(* IEC 61131-3 sources: daoli-st-library/DL_Device (part 3) *)

(* ---- FB_DL_HydraulicPowerUnit.st ---- *)
(*==============================================================================
 * 组件名称 (Component)  : FB_DL_HydraulicPowerUnit
 * 所属子库 (Sublibrary) : DL_Device
 * 当前版本 (Version)    : 1.0.0
 * 兼容性   (Platform)   : CODESYS 3.5+ / TwinCAT 3 / 汇川 InoProShop / 施耐德 Machine Expert
 *                         仅依赖 Standard.library（TON / R_TRIG），零厂商私有库
 * 功能描述 (Function)   : 液压动力单元（HPU）顺控：bStart 上升沿先查油温/油位
 *                         联锁（先于电机判据，规格指定），通过后启动电机升压；
 *                         压力达 fPressSwMpa 开卸荷阀，压力回落至 (fPressSwMpa
 *                         − 0.5 MPa) 关卸荷阀（±0.5 MPa 回差顺控，规格指定）；
 *                         电机启停切换设最小间隔互锁 tMinSw（切换后 tMinSw 内
 *                         禁再次切换）。运行中油温超限/油位低于下限/压力非有限
 *                         → 停电机锁存故障（安全侧优先）。
 * 接口     (Interface)  : 输入 bStart 启动命令（上升沿触发，FALSE 停机）、fPressMpa
 *                         压力实测 [MPa]、fOilTempC 油温实测 [℃]、fOilLevelPct
 *                         油位实测 [%]、fPressSwMpa 卸荷切换阈（域 > 0.5）、
 *                         fTempMaxC 油温联锁上限（域 > 0）、fLvlMinPct 油位联锁
 *                         下限（域 > 0 且 < 100）、tMinSw 电机切换最小间隔、
 *                         bReset 复位；输出 bMotor 电机命令、bUnload 卸荷阀
 *                         命令、ePhase 五态相位、eErrCode 错误码、bError 故障
 *                         标志。
 * 边界     (Boundary)   : ① **属主边界（写死）：本件只出电机/卸荷阀命令，不驱动
 *                         接触器/阀线圈本体**；执行器驱动归 IO 映射层（DOL 电机
 *                         包装归 `FB_DL_DolMotor`）。
 *                         ② 五态 CASE + ELSE 兜底（R6）；tonMinSw IN 挂切换
 *                         互锁窗本身（切换后置互锁、到时解除），三 TON 两沿段 0
 *                         无条件调用（R7）。
 *                         ③ 联锁先于电机判据：启动沿先查油温/油位，联锁不过
 *                         不入启动相并置信息码 eInterlock（不锁存故障，联锁
 *                         为常态门槛）；运行中联锁破约才锁存故障 eTempHigh/
 *                         eLvlLow（归因唯一，R190）。
 *                         ④ 回差口径：开阀阈 fPressSwMpa，关阀阈 fPressSwMpa
 *                         − DL_HPU_DBAND(0.5 MPa)，组态闸保证 fPressSwMpa >
 *                         0.5（关阀阈恒正）。
 *                         ⑤ 电机切换互锁：每次 bMotor 电平变化后 _bSwBlock 置
 *                         位，tonMinSw 到时解除；互锁期内启动/停止命令一律
 *                         拒绝（拒动安全侧）。
 *                         ⑥ 压力非有限（R79 双判）运行中 → 停电机锁存
 *                         ePressBad（不可判即安全侧停机）。
 *                         ⑦ 零全局耦合（无 GVL / VAR_EXTERNAL / 物理地址）。
 * 分工声明 (Scope)      : 与 `FB_DL_DolMotor` 分工：电机直启包装归那件、HPU 工艺
 *                         顺控归本件；与 `FB_DL_MinOnOffGuard` 分工：通用最小
 *                         启停保护归那件，本件互锁为切换间隔专用语义。
 * 来源标签 (Source Tag) : 自研线（卸荷回差顺控为公开液压系统控制实践 clean-room）
 * 码表     (Codes)      : 本件不占用任何全局数字码位。出口为 BOOL 命令组 +
 *                         ENUM 相位/错误码；数字码位待主控收口阶段统一派号。
 * 红线自检 (Redline)    : R1 ✓ 零 GVL/VAR_EXTERNAL ｜ R2 ✓ 零 %I/%Q/%M ｜ R3 ✓ 纯 IEC 61131-3
 *                         R4 ✓ 联锁前置 + 回差 + 切换互锁 + 非有限安全停机
 *                         ｜ R5 ✓ 声明逐行同行双语注释
 *                         R6 ✓ 五态 CASE 含 ELSE ｜ R7 ✓ 三 TON 两 R_TRIG 段 0 无条件刷新
 * 修订历史 (Revision)   : 2026-11-20  v1.0.0  R50 首版（批次 4 · 序号 18）
 * 验收向量 (Acceptance) : ① 油位 25%（下限 30%）时启动沿 → 不入启动相，
 *                         eErrCode=eInterlock，bMotor=FALSE；② 正常启动，
 *                         压力升至 16.2 MPa（阈 16.0）→ bUnload=TRUE；回落至
 *                         15.4 MPa（< 16.0−0.5=15.5）→ bUnload=FALSE；③ 运行
 *                         中油温 65 ℃（上限 60）→ 停电机锁存 eTempHigh；
 *                         ④ 停机后 2s 内再启动（tMinSw=10S）→ 拒动（互锁）。
 *==============================================================================*)

(*-----------------------------------------------------------------------------
 * 枚举: E_DL_HpuPhase（HPU 相位，全库唯一属主本文件）
 *----------------------------------------------------------------------------*)
TYPE E_DL_HpuPhase :
(
    eIdle     := 0,   // 待机（电机停） / Idle, motor off
    eRunning  := 10,  // 升压/运行（电机开，卸荷阀按回差裁决） / Running, unloading by hysteresis
    eFault    := 90   // 故障（等复位） / Fault, awaiting reset
);
END_TYPE

(*-----------------------------------------------------------------------------
 * 枚举: E_DL_HpuErr（错误码；信息级不置 bError，故障级恒伴 bError=TRUE）
 *----------------------------------------------------------------------------*)
TYPE E_DL_HpuErr :
(
    eOk        := 0,   // 正常 / Normal
    eInterlock := 1,   // 信息级：启动被油温/油位联锁拒绝（常态门槛） / Info: start rejected by interlock
    eCfgBad    := 2,   // 故障级：组态非法（阈值/时间域） / Fault: illegal configuration
    eTempHigh  := 3,   // 故障级：运行中油温超限（停电机锁存） / Fault: oil temp high in run
    eLvlLow    := 4,   // 故障级：运行中油位低于下限（停电机锁存） / Fault: oil level low in run
    ePressBad  := 5    // 故障级：压力非有限（安全侧停机锁存） / Fault: pressure non-finite, safe stop
);
END_TYPE

FUNCTION_BLOCK FB_DL_HydraulicPowerUnit
VAR_INPUT
    bStart     : BOOL := FALSE;       // 启动命令（上升沿触发，FALSE 停机请求） [-] / Start command, rising edge triggered
    fPressMpa  : LREAL := 0.0;        // 压力实测 [MPa] / Pressure measurement [MPa]
    fOilTempC  : LREAL := 25.0;       // 油温实测 [℃] / Oil temperature [degC]
    fOilLevelPct: LREAL := 80.0;      // 油位实测 [%] / Oil level [percent]
    fPressSwMpa: LREAL := 16.0;       // 卸荷切换阈（开阀），域 > 0.5 [MPa] / Unload switch threshold
    fTempMaxC  : LREAL := 60.0;       // 油温联锁上限，域 > 0 [℃] / Oil temp interlock ceiling
    fLvlMinPct : LREAL := 30.0;       // 油位联锁下限，域 > 0 且 < 100 [%] / Oil level interlock floor
    tMinSw     : TIME := T#10S;       // 电机切换最小间隔，域 > T#0S [ms] / Minimum motor switch interval
    bReset     : BOOL := FALSE;       // 复位，上升沿清故障锁存（须 bStart=FALSE） [-] / Reset, clears latches when not started
END_VAR
VAR_OUTPUT
    bMotor   : BOOL;                  // 电机命令出口 [-] / Motor command outlet
    bUnload  : BOOL;                  // 卸荷阀命令出口（TRUE=卸荷） [-] / Unload valve command outlet
    ePhase   : E_DL_HpuPhase;         // 相位出口 [-] / Phase outlet
    eErrCode : E_DL_HpuErr;           // 错误码出口 / Error code outlet
    bError   : BOOL;                  // 故障标志（运行联锁破约锁存） [-] / Error flag, latched
END_VAR
VAR
    _eState   : E_DL_HpuPhase := E_DL_HpuPhase.eIdle;   // 内部相（CASE 唯一写入目标） / Internal phase
    _bMot     : BOOL := FALSE;        // 电机命令内部单源（出口同源） / Motor command internal source
    _bUnload  : BOOL := FALSE;        // 卸荷阀内部单源 / Unload valve internal source
    _bFault   : BOOL;                 // 运行故障锁存位（解除沿 = 非启动态 ∧ bReset 上升沿） / Latched run fault bit
    _bCfgBad  : BOOL;                 // 组态非法当拍量 [-] / Illegal configuration
    _bCfgLatch: BOOL;                 // 组态故障锁存位（解除沿 = 非启动态 ∧ bReset 上升沿，与 _bFault 同口径） / Latched config fault
    _bSwBlock : BOOL := FALSE;        // 切换互锁位（切换后置位，tonMinSw 到时解除） / Switch interlock bit
    _bMotPrev : BOOL := FALSE;        // 上拍电机命令快照（切换检测源） / Motor command snapshot
    _bInterlock: BOOL;                // 启动联锁拒绝当拍量（信息级） [-] / Start interlock rejection this scan
    _bNonFin  : BOOL;                 // 压力非有限当拍量 [-] / Pressure non-finite this scan
    _eCause   : E_DL_HpuErr := E_DL_HpuErr.eOk;   // 故障成因锁存（入相时归因，回放不重推断，R189/R190） / Latched fault cause
    rtReset   : R_TRIG;               // 复位沿实例，段 0 无条件调用 / Reset edge instance
    rtStart   : R_TRIG;               // 启动沿实例，段 0 无条件调用 / Start edge instance
    tonMinSw  : TON;                  // 切换互锁窗 TON，段 0 无条件调用（R145：IN 挂互锁位本身） / Switch interlock TON
END_VAR
VAR CONSTANT
    DL_HPU_DBAND : LREAL := 0.5;      // 卸荷回差（关阀阈 = 开阀阈 − 0.5 MPa），规格指定 [MPa] / Unload hysteresis band
    DL_HPU_ZERO  : LREAL := 0.0;      // 判零基准 [MPa] / Zero base
END_VAR

(* —— 段 0：非有限判 + 组态闸 + 三 TON 两沿无条件刷新 —— *)
_bNonFin := (fPressMpa <> fPressMpa) OR ((fPressMpa - fPressMpa) <> DL_HPU_ZERO);   // 压力非有限（R79 双判） / Pressure non-finite
_bCfgBad := (fPressSwMpa <= DL_HPU_DBAND) OR (fTempMaxC <= DL_HPU_ZERO)
         OR (fLvlMinPct <= DL_HPU_ZERO) OR (fLvlMinPct >= 100.0)
         OR (tMinSw <= T#0S);       // 组态域闸（关阀阈恒正保证 + 联锁域 + 互锁窗） / Configuration gate
rtReset(CLK := bReset);             // 复位沿，每拍必调 / Reset edge, every scan
rtStart(CLK := bStart);             // 启动沿，每拍必调 / Start edge, every scan
tonMinSw(IN := _bSwBlock, PT := tMinSw);   // 切换互锁窗（互锁位置位才计时，到时解除） / Switch interlock window

(* —— 段 1：复位沿（须未启动才清锁存；运行中复位无效，安全侧） —— *)
IF rtReset.Q AND (NOT bStart) THEN
    _bFault := FALSE;               // 清运行故障锁存（可达解除路径：停机后复位沿） / Clear run fault
    _bCfgLatch := FALSE;            // 清组态锁存 / Clear config latch
    _eCause := E_DL_HpuErr.eOk;     // 清成因锁存 / Clear cause latch
    _eState := E_DL_HpuPhase.eIdle; // 回待机 / Back to idle
END_IF
IF _bCfgBad AND (NOT _bCfgLatch) THEN
    _bCfgLatch := TRUE;             // 锁存 / Latch
END_IF

(* —— 段 2：电机命令切换检测（电平变化置互锁位；tonMinSw 到时解除） —— *)
IF _bMot <> _bMotPrev THEN
    _bSwBlock := TRUE;              // 切换发生：置互锁（规格⑤） / Switch occurred: engage interlock
END_IF
_bMotPrev := _bMot;                 // 快照（本拍末语义，下一拍比较） / Snapshot for next scan
IF tonMinSw.Q THEN
    _bSwBlock := FALSE;             // 互锁窗到：解除 / Interlock elapsed: release
END_IF

(* —— 段 3：启动联锁判据（先于电机判据，规格③；常态门槛不锁存） —— *)
_bInterlock := (fOilTempC > fTempMaxC) OR (fOilLevelPct < fLvlMinPct);   // 油温/油位联锁 / Oil temp/level interlock

(* —— 段 4：五态顺控（组态/故障期冻结推进；bStart=FALSE 停机优先） —— *)
IF (NOT bStart) OR _bCfgLatch THEN
    _bMot := FALSE;                 // 停机/组态安全侧：电机停 / Stopped or config-safe: motor off
    _bUnload := FALSE;              // 卸荷阀关 / Unload closed
    IF NOT _bFault THEN
        _eState := E_DL_HpuPhase.eIdle;   // 无故障回待机（故障相驻留待复位） / Idle unless fault latched
    END_IF
ELSIF (NOT _bFault) THEN
    CASE _eState OF

    E_DL_HpuPhase.eIdle:
        IF rtStart.Q AND (NOT _bSwBlock) THEN
            IF _bInterlock THEN
                _eState := E_DL_HpuPhase.eIdle;   // 联锁不过：拒绝启动（信息码见段 6，R191 声明） / Interlock rejected
            ELSE
                _bMot := TRUE;    // 电机启动 / Motor on
                _eState := E_DL_HpuPhase.eRunning;   // 入运行相 / Enter running
            END_IF
        END_IF

    E_DL_HpuPhase.eRunning:
        (* 运行中联锁破约/压力非有限 → 停电机锁存故障（安全侧优先，规格⑥） *)
        IF fOilTempC > fTempMaxC THEN
            _bMot := FALSE;       // 停电机 / Motor off
            _bFault := TRUE;      // 锁存 / Latch
            _eCause := E_DL_HpuErr.eTempHigh;   // 入相归因：油温超限 / Cause at entry: temp high
            _eState := E_DL_HpuPhase.eFault;   // 入故障相 / Enter fault
        ELSIF fOilLevelPct < fLvlMinPct THEN
            _bMot := FALSE;       // 停电机 / Motor off
            _bFault := TRUE;      // 锁存 / Latch
            _eCause := E_DL_HpuErr.eLvlLow;     // 入相归因：油位低 / Cause at entry: level low
            _eState := E_DL_HpuPhase.eFault;   // 入故障相 / Enter fault
        ELSIF _bNonFin THEN
            _bMot := FALSE;       // 压力不可判：安全侧停机（规格⑥） / Pressure unjudgeable: safe stop
            _bFault := TRUE;      // 锁存 / Latch
            _eCause := E_DL_HpuErr.ePressBad;   // 入相归因：压力非有限 / Cause at entry: pressure non-finite
            _eState := E_DL_HpuPhase.eFault;   // 入故障相 / Enter fault
        ELSE
            (* 卸荷回差顺控（±0.5 MPa，规格④）：开阀阈 / 关阀阈容差比较 *)
            IF (NOT _bUnload) AND (fPressMpa >= fPressSwMpa) THEN
                _bUnload := TRUE;   // 达开阀阈：卸荷 / At open threshold: unload
            ELSIF _bUnload AND (fPressMpa <= (fPressSwMpa - DL_HPU_DBAND)) THEN
                _bUnload := FALSE;  // 回落至关阀阈：加载 / Back to close threshold: load
            END_IF
        END_IF

    E_DL_HpuPhase.eFault:
        ;                         // 故障相驻留（由复位沿迁出链处理） / Held by reset chain

    ELSE
        _bMot := FALSE;           // 非法相位兜底：电机安全侧停 / Illegal phase: safe stop
        _bUnload := FALSE;        // 卸荷阀关 / Unload closed
        _bFault := TRUE;          // 锁存（R45 配对见段 6） / Latch
        _eCause := E_DL_HpuErr.eCfgBad;   // 兜底归因：按组态级回放 / Fallback cause: config level
        _eState := E_DL_HpuPhase.eFault;   // 强拉故障相 / Force fault phase

    END_CASE
END_IF

(* —— 段 5：出口单点映射（名实双出口同源，R191） —— *)
bMotor := _bMot;                  // 电机命令出口 / Motor command outlet
bUnload := _bUnload;              // 卸荷阀命令出口 / Unload command outlet
ePhase := _eState;                // 相位出口 / Phase outlet
IF _bCfgLatch THEN
    bError := TRUE;               // 故障标志（R45 配对） / Error flag
    eErrCode := E_DL_HpuErr.eCfgBad;   // 组态级码 / Config fault code
ELSIF _bFault THEN
    bError := TRUE;               // 故障标志 / Error flag
    eErrCode := _eCause;          // 成因锁存回放（禁故障相当拍重推断，R189） / Cause latch replay
ELSE
    bError := FALSE;              // 无故障级条件 / No fault
    IF _bInterlock AND rtStart.Q AND (NOT _bSwBlock) THEN
        eErrCode := E_DL_HpuErr.eInterlock;   // 信息级：启动联锁拒绝（当拍） / Info: start rejected
    ELSE
        eErrCode := E_DL_HpuErr.eOk;          // 正常 / Normal
    END_IF
END_IF

END_FUNCTION_BLOCK

(* ---- FB_DL_LevelRadarValidate.st ---- *)
(*==============================================================================
 * 组件名称 (Component)  : FB_DL_LevelRadarValidate
 * 溯源说明 (Provenance): 道莅 clean-room 防御性实现（IEC 61131-3 纯净实现，闭源文档仅借语义，零代码行）
 * 所属子库 (Sublibrary) : DL_Device / SignalQuality
 * 当前版本 (Version)    : 1.0.0
 * 兼容性   (Platform)   : CODESYS 3.5 / TwinCAT 3 / 汇川 InoProShop / 施耐德
 *                         Machine Expert；纯 IEC 61131-3（第 3 版），仅用
 *                         Standard.library 的 TON / ABS / LIMIT / TIME_TO_REAL
 * 组件分类 (Category)   : 功能块（FUNCTION_BLOCK）· 雷达液位回波可信度仲裁
 * 功能一句话 (Summary)  : 用回波置信度、信噪比、量程、变化率四条判据仲裁雷达液位
 *                         是否可信，不可信时保持末次可信值并给出四位掩码。
 *
 * 本件存在的意义 (Why this unit exists)
 *   雷达液位最典型的失效不是「没读数」，而是**读数看着很正常但其实是假回波**
 *   （搅动液面、泡沫、罐壁多重反射）。一旦假回波进了联锁或计量，结果是
 *   抽空泵或溢出。I_DL_AnalogSensor 只管 4~20 mA 的质量位，解不了回波域；
 *   本件补的正是「回波可信度」这一层。
 *
 * 四判据同拍评估（**不早退**，全部写进掩码）
 *   位 1 置信度低 : fQuality < fQualityMin
 *   位 2 信噪比低 : fSnr < fSnrMin
 *   位 4 超量程   : fLevel < 0 或 fLevel > fSpan
 *   位 8 变化率跳变: |fLevel − 末次可信值| / 采样周期 > fRateLimit
 *   四条同时评估、同时写进掩码——现场要的是「一次看全四条」，早退只会让人
 *   改一条跑一次。bTrusted = (uSuspectMask = 0) 即时给出（联锁看即时值，
 *   不能等确认窗）。
 *
 * 状态抖动抑制 (Anti-flicker)
 *   进入不可信是**即时**的（假回波必须立刻挡住），恢复可信要 mask 全零
 *   持续 tConfirm 才生效。这是一条不对称的滞回：宁可晚一点恢复，也不让
 *   读数在临界回波上反复跳。
 *
 * 边界安全 (Boundary)
 *   ① fSpan <= 0、门限非法或采样周期 <= 0 → 故障 0345、bValid = FALSE；
 *   ② 任一输入非有限 → 故障 0346，**本次不更新 fLevelOut**（R42：跨拍取值必须
 *      本拍复验，坏值绝不进联锁）；
 *   ③ 超量程只置掩码位，不按可信值发布；
 *   ④ 初始无历史可信值 → fLevelOut := 0 且 bValid := FALSE，**绝不把 0 m 当可信
 *      液位发布**（R43 家族：保持值必须夹进有效域并标记不可用）；
 *   ⑤ 失能 → bTrusted := FALSE、eHealth := eUnknown，fLevelOut 保持（供趋势）；
 *   ⑥ 采样周期由 tSample 引脚注入，**禁读系统时钟**；
 *   ⑦ CASE 落 ELSE 置 0347 并回 eFault。
 *
 * 错误码    : 16#0003_0178 质量指标低于门限，保持末次可信值——信息级，正常防御
 *             16#0003_0179 变化率跳变，单拍剔除——信息级，正常防御
 *             16#0003_0345 量程/门限/采样周期参数非法——故障级，bValid = FALSE
 *             16#0003_0346 输入非有限，不更新发布值——故障级
 *             16#0003_0347 状态机落 ELSE 兜底（非法状态）——故障级，回 eFault
 * 码位总账  : 16#0003_0178 用 / 16#0003_0179 用 ｜ 16#0003_0345 用 / 16#0003_0346 用 / 16#0003_0347 用
 * 状态机    : E_DL_RadarState（eIdle / eTrusted / eSuspect / eFault），CASE 含 ELSE 兜底，
 *             ELSE 置 16#0003_0347 并回 eFault；失能无条件回 eIdle
 * 采样约定  : 每任务周期调用一次；变化率判据用 tSample 引脚换算，不读系统时钟
 * 依赖说明  : 仅 Standard.library；健康出口引用 E_DL_Ne107Status（引用不重声明，R70③）
 * 验收向量  : V1 液位 5.00 m、置信度 80 %、信噪比 20 dB、量程 10 m、上拍可信 4.98
 *               → bTrusted = TRUE，uSuspectMask = 0，fLevelOut = 5.00，eHealth = eOk
 *             V2 置信度 20 %（< 40）→ 掩码位 1，bTrusted = FALSE，fLevelOut 保持 4.98，
 *                eErr = 0178，eHealth = eCheckFunction（保持主向量）
 *             V3 液位 12.0 m（> 量程 10），置信度与信噪比都好 → 掩码位 4，
 *                不按可信值发布（超量程主向量）
 *             V4 上拍可信 1.00 m，本拍 6.00 m、tSample 1 s、fRateLimit 0.5 m/s
 *                → 掩码位 8 + 位 1/2 若同时成立全部置位，eErr 优先级见段 9（跳变主向量）
 *             V5 冷启动首拍（无历史可信值）且本拍不可信 → fLevelOut = 0 且 bValid = FALSE
 *                （R43 主向量：0 m 绝不发布为可信液位）
 *             V6 fLevel = NaN → 0346，fLevelOut 不更新（坏值不进联锁主向量）
 *             V7 fSpan = 0 → 0345，bValid = FALSE
 *             V8 恢复：mask 全零但未满 tConfirm → 仍 eSuspect；满窗 → eTrusted（滞回主向量）
 * 红线自检  : 全局变量声明零使用 / 外部变量访问零使用 / 物理地址零使用 ｜ 纯 IEC 61131-3 ｜ 除零前置
 *             闸（tSample 恒 > 0 且商前显式判据）｜ 浮点只用大小与容差比较 ｜ 无循环
 *             ｜ 全变量双语同行注释 ｜ ENUM + CASE 含 ELSE ｜ TON 在主体前部无条件
 *             刷新 ｜ 掩码与阈值常量化，无魔法数
 * 修订历史  : 2026-11-16  v1.0.0  首版入库（R22 · 批 3 · 设备信号质量）
 *============================================================================*)

(*-----------------------------------------------------------------------------
 * 枚举: E_DL_RadarState（归属本功能块，同文件发布，全库唯一定义）
 * 含义: 回波仲裁相位。0 起步长 10。
 *-----------------------------------------------------------------------------*)
TYPE E_DL_RadarState :
(
    eIdle    := 0,     // 待机：未使能或参数非法 / Idle, disabled or illegal parameters
    eTrusted := 10,    // 可信：四条判据全部通过 / Trusted, all four criteria pass
    eSuspect := 20,    // 存疑：至少一条判据失败，发布值保持 / Suspect, at least one criterion failed
    eFault   := 99     // 故障：参数非法或输入非有限 / Fault, illegal parameter or non-finite input
);
END_TYPE

FUNCTION_BLOCK FB_DL_LevelRadarValidate
VAR_INPUT
    fLevel       : REAL;                       // 雷达测得液位 [m] / radar measured level [m]
    fQuality     : REAL;                       // 回波置信度 [%]，范围 0~100 / echo confidence [%], range 0~100
    fSnr         : REAL;                       // 回波信噪比 [dB] / echo signal to noise ratio [dB]
    fSpan        : REAL := 10.0;               // 量程上限 [m]，须 > 0 / span ceiling [m], must be > 0
    fQualityMin  : REAL := 40.0;               // 置信度门限 [%]，范围 0~100 / confidence threshold [%], range 0~100
    fSnrMin      : REAL := 10.0;               // 信噪比门限 [dB]，须 >= 0 / signal to noise threshold [dB], must be >= 0
    fRateLimit   : REAL := 0.5;                // 液位变化率上限 [m/s]，须 > 0 / level rate ceiling [m/s], must be > 0
    tConfirm     : TIME := T#10S;              // 恢复可信确认时间 [ms] / recovery confirm time [ms]
    tSample      : TIME := T#1S;               // 采样周期 [ms]，变化率换算用 / sample period [ms], used by the rate test
    bEnable      : BOOL;                       // 使能 / enable
END_VAR
VAR_OUTPUT
    fLevelOut    : REAL;                       // 发布值：可信则实时值，否则末次可信值 [m] / published level [m]
    bTrusted     : BOOL;                       // 本拍回波可信 / this scan's echo is trusted
    uSuspectMask : WORD;                       // 存疑位掩码：1 置信度 / 2 信噪比 / 4 超量程 / 8 跳变
    eHealth      : E_DL_Ne107Status;           // NE107 健康分级（引用唯一属主） / NE107 health status
    eErr         : UDINT;                      // 错误码，0 表示无错 / error code, 0 means no error
    bError       : BOOL;                       // 故障级标志，仅故障级错误置位 / fault-class flag, set only on fault-level codes
    bValid       : BOOL;                       // 发布值可用标志 / published value usable flag
END_VAR
VAR
    fbTrust      : TON;                        // 恢复可信确认窗，段 6 无条件刷新 [ms] / recovery confirm window
    _eState      : E_DL_RadarState := E_DL_RadarState.eIdle; // 当前相位 / current phase
    _bInit       : BOOL := FALSE;              // 首扫标志，初值 FALSE 取非判定 / first-scan flag, tested negated
    _bParamBad   : BOOL;                       // 参数非法标志 / illegal parameter flag
    _bFiniteBad  : BOOL;                       // 输入非有限标志 / non-finite input flag
    _bIllegal    : BOOL;                       // 非法状态标志 / illegal state flag
    _bHaveTrusted : BOOL;                      // 是否已有历史可信值 / whether a trusted value exists
    _bBrkTrust   : BOOL;                       // 恢复确认计时器断输入一拍 / recovery timer one-scan break
    _bBadQuality : BOOL;                       // 置信度不足 / confidence too low
    _bBadSnr     : BOOL;                       // 信噪比不足 / signal to noise too low
    _bBadSpan    : BOOL;                       // 超量程 / out of span
    _bBadRate    : BOOL;                       // 变化率跳变 / rate jump
    _tConfirmUse : TIME := T#10S;              // 生效确认时间 [ms]，已钳位 / effective confirm time, clamped
    _fDtSec      : REAL := 1.0;                // 生效采样周期 [s] / effective sample period [s]
    _fLastTrusted : REAL;                      // 末次可信液位 [m] / last trusted level [m]
    _fOutHeld    : REAL;                       // 发布值保持量 [m] / held published level [m]
    _fRate       : REAL;                       // 本拍变化率 [m/s] / level rate of this scan [m/s]
    _wMask       : WORD;                       // 本拍掩码暂存 / mask staging of this scan
END_VAR
VAR CONSTANT
    DL_VAL_LIM     : REAL := 1.0E6;            // 有限性判定的绝对值上限 [无量纲] / finiteness ceiling
    DL_LEVEL_MIN   : REAL := 0.0;              // 液位物理下限 [m] / level physical floor [m]
    DL_QUAL_MAX    : REAL := 100.0;            // 置信度上限 [%] / confidence ceiling [%]
    DL_QUAL_MIN    : REAL := 0.0;              // 置信度下限 [%] / confidence floor [%]
    DL_SNR_MIN     : REAL := 0.0;              // 信噪比下限 [dB] / signal to noise floor [dB]
    DL_SPAN_MIN    : REAL := 0.0;              // 量程下限 [m]，须严格大于 / span floor [m], strictly greater
    DL_RATE_MIN    : REAL := 0.0;              // 变化率上限下限 [m/s]，须严格大于 / rate floor [m/s], strictly greater
    DL_MS_PER_S    : REAL := 1000.0;           // 毫秒与秒的换算系数 [ms/s] / milliseconds per second
    DL_ONE_SEC     : REAL := 1.0;              // 一秒的兜底值 [s]，采样周期非法时使用 / one second fallback [s]
    DL_CONF_MAX_MS : DINT := 3600000;          // 确认时间上限 [ms]，一小时 / confirm time ceiling, one hour
    DL_TIME_ZERO   : TIME := T#0MS;            // 时间零值基准 [ms] / time zero reference
    DL_MASK_QUAL   : WORD := 16#0001;          // 掩码位 1：置信度低 / mask bit one, low confidence
    DL_MASK_SNR    : WORD := 16#0002;          // 掩码位 2：信噪比低 / mask bit two, low signal to noise
    DL_MASK_SPAN   : WORD := 16#0004;          // 掩码位 4：超量程 / mask bit four, out of span
    DL_MASK_RATE   : WORD := 16#0008;          // 掩码位 8：变化率跳变 / mask bit eight, rate jump
    DL_MASK_NONE   : WORD := 16#0000;          // 无存疑 / no suspicion
END_VAR

(*------------------------------------------------------------------------------
 * 段 1｜每拍预置（发布值与保持量在段 8 单点写入）
 *      Per-scan presets, the published value is written only in segment eight
 *-----------------------------------------------------------------------------*)
eErr         := 16#0000_0000;                  // 错误码每拍重算 / error code recomputed every scan
bError       := FALSE;                         // 故障标志每拍重算 / fault flag recomputed every scan
bValid       := FALSE;                         // 可用标志每拍重算 / usable flag recomputed every scan
bTrusted     := FALSE;                         // 可信标志每拍重算 / trusted flag recomputed
uSuspectMask := DL_MASK_NONE;                  // 掩码清零 / mask cleared
_bParamBad   := FALSE;                         // 参数非法标志预清零 / parameter flag pre-cleared
_bFiniteBad  := FALSE;                         // 非有限标志预清零 / non-finite flag pre-cleared
_bIllegal    := FALSE;                         // 非法状态标志预清零 / illegal state flag pre-cleared
_bBadQuality := FALSE;                         // 置信度判据预置 FALSE / confidence criterion preset FALSE
_bBadSnr     := FALSE;                         // 信噪比判据预置 FALSE / snr criterion preset FALSE
_bBadSpan    := FALSE;                         // 量程判据预置 FALSE / span criterion preset FALSE
_bBadRate    := FALSE;                         // 变化率判据预置 FALSE / rate criterion preset FALSE
_wMask       := DL_MASK_NONE;                  // 掩码暂存清零 / mask staging cleared
_fRate       := 0.0;                           // 变化率预置 0 [m/s] / rate preset to zero

(*------------------------------------------------------------------------------
 * 段 2｜首扫初始化（**无历史可信值**：0 m 不是液位，是「还没有数据」）
 *      First-scan initialisation, no trusted value exists yet
 *-----------------------------------------------------------------------------*)
IF NOT _bInit THEN
    _eState       := E_DL_RadarState.eIdle;    // 相位待机 / phase idle
    _fLastTrusted := 0.0;                      // 末次可信值 0 [m] / last trusted level zero
    _fOutHeld     := 0.0;                      // 发布值保持量 0 [m] / held published value zero
    _bHaveTrusted := FALSE;                    // 尚无历史可信值 / no trusted value yet
    _bBrkTrust    := TRUE;                     // 恢复确认窗从零开始 / recovery window starts from zero
    _bInit        := TRUE;                     // 首扫只做一次 / the first scan runs once
END_IF

(*------------------------------------------------------------------------------
 * 段 3｜参数闸门（量程、四条门限与采样周期；除零前置闸在采样周期处）
 *      Parameter gate, the sample period guard also protects the rate division
 *-----------------------------------------------------------------------------*)
IF (fSpan <> fSpan) OR (ABS(fSpan) > DL_VAL_LIM) OR (fSpan <= DL_SPAN_MIN) THEN
    _bParamBad := TRUE;                        // 量程非法 / span illegal
END_IF
IF (fQualityMin <> fQualityMin) OR (fQualityMin < DL_QUAL_MIN) OR (fQualityMin > DL_QUAL_MAX) THEN
    _bParamBad := TRUE;                        // 置信度门限非法 / confidence threshold illegal
END_IF
IF (fSnrMin <> fSnrMin) OR (fSnrMin < DL_SNR_MIN) OR (ABS(fSnrMin) > DL_VAL_LIM) THEN
    _bParamBad := TRUE;                        // 信噪比门限非法 / snr threshold illegal
END_IF
IF (fRateLimit <> fRateLimit) OR (ABS(fRateLimit) > DL_VAL_LIM) OR (fRateLimit <= DL_RATE_MIN) THEN
    _bParamBad := TRUE;                        // 变化率上限非法 / rate ceiling illegal
END_IF

_tConfirmUse := tConfirm;                      // 确认时间直取引脚 [ms] / confirm time from the pin
IF TIME_TO_DINT(_tConfirmUse) > DL_CONF_MAX_MS THEN
    _tConfirmUse := DINT_TO_TIME(DL_CONF_MAX_MS); // 超上限钳位（无专用码位，R90 不新开码） / clamped
END_IF
IF TIME_TO_DINT(tSample) <= 0 THEN
    _bParamBad := TRUE;                        // 采样周期非正：变化率判据无意义 / non-positive sample period
    _fDtSec    := DL_ONE_SEC;                  // 兜底 1 s，防后续除零 / fallback to one second, no division by zero
ELSE
    _fDtSec := TIME_TO_REAL(tSample) / DL_MS_PER_S; // 采样周期换算为秒 [s] / sample period in seconds
END_IF
IF _fDtSec <= DL_RATE_MIN THEN
    _fDtSec := DL_ONE_SEC;                     // 结构性兜底：商恒 > 0，仍显式判一次 / explicit fallback, defense in depth
END_IF

(*------------------------------------------------------------------------------
 * 段 4｜输入有限性（区间判据同时拦 NaN 与 ±Inf）
 *      Input finiteness, the interval test catches NaN and infinity
 *-----------------------------------------------------------------------------*)
IF (fLevel < -DL_VAL_LIM) OR (fLevel > DL_VAL_LIM) THEN
    _bFiniteBad := TRUE;                       // 液位非有限 / level non-finite
END_IF
IF (fQuality < -DL_VAL_LIM) OR (fQuality > DL_VAL_LIM) THEN
    _bFiniteBad := TRUE;                       // 置信度非有限 / confidence non-finite
END_IF
IF (fSnr < -DL_VAL_LIM) OR (fSnr > DL_VAL_LIM) THEN
    _bFiniteBad := TRUE;                       // 信噪比非有限 / snr non-finite
END_IF

(*------------------------------------------------------------------------------
 * 段 5｜四条判据同拍评估（不早退：全部写进掩码，便于现场一次改全）
 *      All four criteria evaluated in the same scan, no early exit
 *-----------------------------------------------------------------------------*)
IF (NOT _bFiniteBad) AND (NOT _bParamBad) THEN
    _bBadQuality := (fQuality < fQualityMin);  // 判据 1：置信度低 / criterion one, low confidence
    _bBadSnr     := (fSnr < fSnrMin);          // 判据 2：信噪比低 / criterion two, low snr
    _bBadSpan    := (fLevel < DL_LEVEL_MIN) OR (fLevel > fSpan); // 判据 3：超量程 / criterion three, out of span

    IF _bHaveTrusted THEN
        _fRate := ABS(fLevel - _fLastTrusted) / _fDtSec; // 变化率 [m/s]，除数恒 > 0 / rate, the divisor is always positive
    ELSE
        _fRate := 0.0;                         // 无历史可信值：不判跳变（首次读数无基准） / no baseline yet
    END_IF
    _bBadRate := (_fRate > fRateLimit);        // 判据 4：变化率跳变 / criterion four, rate jump

    IF _bBadQuality THEN
        _wMask := _wMask OR DL_MASK_QUAL;      // 置置信度位 / set the confidence bit
    END_IF
    IF _bBadSnr THEN
        _wMask := _wMask OR DL_MASK_SNR;       // 置信噪比位 / set the snr bit
    END_IF
    IF _bBadSpan THEN
        _wMask := _wMask OR DL_MASK_SPAN;      // 置超量程位 / set the span bit
    END_IF
    IF _bBadRate THEN
        _wMask := _wMask OR DL_MASK_RATE;      // 置跳变位 / set the rate bit
    END_IF
END_IF

(*------------------------------------------------------------------------------
 * 段 6｜恢复确认计时器无条件刷新（进入不可信是即时的，恢复才要确认窗）
 *      Recovery timer refreshed unconditionally, entry is immediate, exit needs the window
 *-----------------------------------------------------------------------------*)
fbTrust(IN := bEnable AND (NOT _bFiniteBad) AND (NOT _bParamBad) AND (_wMask = DL_MASK_NONE)
             AND (NOT _bBrkTrust), PT := _tConfirmUse); // 恢复可信确认窗
_bBrkTrust := FALSE;                           // 断输入拍在调用后自清 / break self-cleared after the call

(*------------------------------------------------------------------------------
 * 段 7｜相位机（进入存疑即时，退出存疑须窗满；不对称滞回）
 *      Phase machine with an asymmetric hysteresis
 *-----------------------------------------------------------------------------*)
CASE _eState OF

    E_DL_RadarState.eIdle:                     // 待机：参数合法且使能即判可信度
        IF _bParamBad OR _bFiniteBad THEN
            _eState := E_DL_RadarState.eFault; // 原因未消失，转故障 / the cause persists
        ELSIF bEnable THEN
            IF _wMask = DL_MASK_NONE THEN
                _eState := E_DL_RadarState.eTrusted; // 首拍即可信 / trusted from the first scan
            ELSE
                _eState := E_DL_RadarState.eSuspect; // 首拍即存疑 / suspect from the first scan
            END_IF
        END_IF

    E_DL_RadarState.eTrusted:                  // 可信：任一判据失败即时转存疑
        IF _bParamBad OR _bFiniteBad THEN
            _eState := E_DL_RadarState.eFault; // 转故障 / go to fault
        ELSIF NOT bEnable THEN
            _eState := E_DL_RadarState.eIdle;  // 失能回待机 / disabled, back to idle
        ELSIF _wMask <> DL_MASK_NONE THEN
            _eState := E_DL_RadarState.eSuspect; // 即时转存疑（假回波必须立刻挡住） / immediate, a false echo must be blocked
            _bBrkTrust := TRUE;                // 恢复窗重启 / the recovery window restarts
        END_IF

    E_DL_RadarState.eSuspect:                  // 存疑：掩码全零且满窗才恢复
        IF _bParamBad OR _bFiniteBad THEN
            _eState := E_DL_RadarState.eFault; // 转故障 / go to fault
        ELSIF NOT bEnable THEN
            _eState := E_DL_RadarState.eIdle;  // 失能回待机 / disabled, back to idle
        ELSIF (_wMask = DL_MASK_NONE) AND fbTrust.Q THEN
            _eState := E_DL_RadarState.eTrusted; // 满窗恢复可信 / recovered after the window
        END_IF

    E_DL_RadarState.eFault:                    // 故障：参数与输入恢复即可回待机
        IF bEnable AND (NOT _bParamBad) AND (NOT _bFiniteBad) THEN
            _eState := E_DL_RadarState.eIdle;  // 原因消失 / the cause is gone
            _bBrkTrust := TRUE;                // 恢复窗重启，避免沿用故障期残留 / the window restarts
        END_IF

    ELSE
        _bIllegal := TRUE;                     // 标记非法状态 / flag the illegal state
        _eState   := E_DL_RadarState.eFault;   // 回故障态 / back to the fault state
END_CASE

(*------------------------------------------------------------------------------
 * 段 8｜发布值单点写入（可信用实时值，否则保持；无历史时 0 且不可用）
 *      Single write point of the published value
 *-----------------------------------------------------------------------------*)
IF (NOT _bFiniteBad) AND (NOT _bParamBad) AND (_wMask = DL_MASK_NONE) THEN
    _fOutHeld     := fLevel;                   // 可信：发布实时值 [m] / trusted, publish the live value
    _fLastTrusted := fLevel;                   // 同步末次可信值 [m] / latch the last trusted value
    _bHaveTrusted := TRUE;                     // 已有历史可信值 / a trusted value now exists
END_IF
(* 不可信拍一律不更新 _fOutHeld：保持末次可信值 / an untrusted scan leaves the held value untouched *)

fLevelOut    := _fOutHeld;                     // 发布值出口 [m] / published value outlet
uSuspectMask := _wMask;                        // 存疑掩码出口 / suspect mask outlet
bTrusted     := ((_wMask = DL_MASK_NONE) AND (NOT _bFiniteBad) AND (NOT _bParamBad) AND bEnable); // 即时可信标志

(*------------------------------------------------------------------------------
 * 段 9｜码位优先级链与健康分级
 *      Code priority chain and health grading
 *-----------------------------------------------------------------------------*)
IF _bIllegal THEN
    eErr   := 16#0003_0347;                    // 故障级：状态机兜底 / fault: state machine fallback
    bError := TRUE;                            // 置故障标志 / raise the fault flag
ELSIF _bParamBad THEN
    eErr   := 16#0003_0345;                    // 故障级：量程/门限/采样周期非法 / fault: span, thresholds or sample period illegal
    bError := TRUE;                            // 置故障标志 / raise the fault flag
ELSIF _bFiniteBad THEN
    eErr   := 16#0003_0346;                    // 故障级：输入非有限，不更新发布值 / fault: non-finite input
    bError := TRUE;                            // 置故障标志 / raise the fault flag
ELSIF _bBadRate THEN
    eErr   := 16#0003_0179;                    // 信息级：变化率跳变，单拍剔除 / informational: rate jump rejected
ELSIF _wMask <> DL_MASK_NONE THEN
    eErr   := 16#0003_0178;                    // 信息级：质量指标低于门限，保持末次可信值 / informational: quality below threshold
END_IF

IF _bParamBad OR _bFiniteBad OR _bIllegal THEN
    eHealth := E_DL_Ne107Status.eFailure;      // 无判定能力：失效 / no verdict capability
ELSIF NOT bEnable THEN
    eHealth := E_DL_Ne107Status.eUnknown;      // 失能：无结论 / disabled, no verdict
ELSIF _wMask <> DL_MASK_NONE THEN
    eHealth := E_DL_Ne107Status.eCheckFunction; // 回波存疑：需检查功能（探头/泡沫/扰动） / suspect echo, check function
ELSE
    eHealth := E_DL_Ne107Status.eOk;           // 回波可信 / trusted echo
END_IF

IF bError THEN
    bValid := FALSE;                           // 故障级：发布值不可用 / fault: unusable
ELSIF NOT bEnable THEN
    bValid := FALSE;                           // 失能：发布值不可用 / disabled: unusable
ELSIF NOT _bHaveTrusted THEN
    bValid := FALSE;                           // 无历史可信值：0 m 绝不作为可信液位发布（R43） / never publish zero as trusted
ELSE
    bValid := TRUE;                            // 发布值可用（存疑时为末次可信值，仍可用） / usable, the held value is still valid
END_IF

END_FUNCTION_BLOCK

(* ---- FB_DL_LoadCellTareDrift.st ---- *)
(*==============================================================================
 * 组件名称 (Component)  : FB_DL_LoadCellTareDrift
 * 所属子库 (Sublibrary) : DL_Device
 * 当前版本 (Version)    : 1.0.0
 * 兼容性   (Platform)   : CODESYS 3.5+ / TwinCAT 3 / 汇川 InoProShop / 施耐德 Machine Expert
 *                         仅依赖 Standard.library（TON / R_TRIG / ABS），零厂商私有库
 * 功能描述 (Function)   : 称重零点漂移监视与去皮闸。
 *                           ① 去皮：bTareCmd 上升沿且**去皮闸放行**时才取当前重量为去皮基准
 *                              fTareRef，并出单拍 bTareDone；闸门未满足则 bTareRejected 且不动基准
 *                              （不"先去了再报错"——那会把错误的零点写进台账）。
 *                           ② 去皮闸三条件同时成立：空载 bNoLoad、|fWeight| 在稳定带
 *                              fTareStableBand 内、且该状态持续 tTareStable（tonStable）。
 *                           ③ 漂移监视：以周期窗 tonObserve（自复位周期窗）为节拍，在窗末取
 *                              当拍重量与去皮基准之差 fDrift，除以窗长（分钟）得漂移速率
 *                              fDriftRate；按 fDriftWarnRate / fDriftAlarmRate 判三级。
 *                              速率判级只在空载时可信（载重下的读数变化是载荷不是漂移），
 *                              故 bNoLoad=FALSE 时维持上一速率不刷新、也不升级告警。
 * 接口     (Interface)  : 输入 fWeight 当前重量、bNoLoad 空载判定（外部给）、fDriftWarnRate /
 *                         fDriftAlarmRate 漂移速率档（单位/分钟）、tObserveWin 观测窗（TIME）、
 *                         fObserveWinMin 同一窗长的分钟数值（REAL，与 tObserveWin 成对给）、
 *                         fTareStableBand 去皮稳定带、tTareStable 去皮稳定时间、bTareCmd 去皮命令、
 *                         bReset 复位；输出 fTareRef 去皮基准、fBaseline 空载基线、fDriftRate 漂移
 *                         速率、eGrade 判级、bTareAllowed 去皮闸状态、bTareDone 去皮完成单拍、
 *                         bTareRejected 去皮被拒、bAlarm 漂移报警锁存、eState / eCause / bError。
 * 边界     (Boundary)   : ① **PT 语义成对声明（R228A 豁免说明的配套要求）**：任何"用 TIME 计时、
 *                         又要用数值参与换算"的地方，一律由调用方**同时**给 TIME 与 REAL 两个
 *                         同义引脚（tObserveWin 与 fObserveWinMin）。本件**不做 TIME→数值转换**，
 *                         从根上避开 TIME_TO_DINT 在各平台单位/可用性差异与"恒假判据"类缺陷。
 *                         调用方必须保证二者一致（同一窗长），不一致属调用方组态错误，本件无法
 *                         在内部交叉校验（那需要 TIME→数值，正是要避开的操作）。
 *                         ② 组态闸：tObserveWin <= T#0S、fObserveWinMin <= DL_LCT_EPS、
 *                         fDriftWarnRate <= 0.0、fDriftAlarmRate <= fDriftWarnRate、
 *                         fTareStableBand <= 0.0、tTareStable < T#0S、任一浮点 NaN → 故障锁存，
 *                         去皮闸强制关闭（宁可不去皮，不可错去皮）。
 *                         ③ 本件**不做温度补偿、不改标定系数**，只做零点漂移监视与去皮闸；
 *                         标定与温度补偿属称重仪表内部职能或上层标定件。
 *                         ④ 三枚 TON/两枚 R_TRIG 段 0 无条件周期刷新；tonObserve 用
 *                         IN := (NOT tonObserve.Q) 自复位形成周期窗（R188 合规写法）。
 *                         ⑤ 故障相与报警锁存迁出唯一路径 = bReset 上升沿（R228B）。
 *                         ⑥ 零全局耦合（无 GVL / 无 VAR_EXTERNAL / 无物理地址）。
 * 分工声明 (Scope)      : 与 `FB_DL_AxisTorqueLimitGuard` 一类力/矩监控件分工——那些判瞬时超限，
 *                         本件判**零点慢漂**（分钟级趋势），时间尺度差三个数量级以上，不可互替。
 * 来源标签 (Source Tag) : T2-2 ◐（开源参考：称重去皮与零点漂移监视参数域，零代码行复制）
 * 解除式   (Release)    : bReset 上升沿 ∧ 组态合法 ∧ 当拍 bNoLoad ∧ 当拍 |fDriftRate| < fDriftWarnRate
 *                         （R240 全当拍量）。自证可满足：重新去皮或载荷卸空即满足，无死锁。
 * 码表     (Codes)      : 本件不占用任何全局数字码位。出口为 ENUM 判级 + BOOL 组（bTareDone /
 *                         bTareRejected / bAlarm / bError）；数字码位待主控收口阶段统一派号。
 * 红线自检 (Redline)    : R1 ✓ 零 GVL/VAR_EXTERNAL ｜ R2 ✓ 零 %I/%Q/%M ｜ R3 ✓ 纯 IEC 61131-3
 *                         R4 ✓ 除零闸 + 阈值几何闸 + 浮点容差 ｜ R5 ✓ 声明逐行同行双语注释
 *                         R6 ✓ ENUM+CASE 含 ELSE ｜ R7 ✓ TON/R_TRIG 段 0 无条件刷新
 * 修订历史 (Revision)   : 2026-11-19  v1.0.0  R46 首版（批次 2 · 序号 9）
 *==============================================================================*)

TYPE E_DL_LctGrade :
(
    eUnknown := 0,    // 尚未测得速率 / Rate not measured yet
    eOk      := 10,   // 漂移在预警带内 / Drift inside the warning band
    eWarn    := 20,   // 漂移达预警档（维护级） / Drift at the warning level
    eAlarm   := 30    // 漂移达报警档（锁存） / Drift at the alarm level, latched
);
END_TYPE

TYPE E_DL_LctState :
(
    eIdle  := 0,    // 首次去皮的等待相 / Awaiting the first tare
    eRun   := 10,   // 漂移监视运行相 / Drift monitoring phase
    eFault := 90    // 组态故障相（去皮闸强制关闭） / Configuration fault, tare gate forced closed
);
END_TYPE

TYPE E_DL_LctCause :
(
    eNone        := 0,   // 无异常 / No anomaly
    eCfgIllegal  := 1,   // 组态非法 / Illegal configuration
    eTareReject  := 2,   // 去皮被拒（未空载/未稳定/超稳定带） / Tare rejected, gate not satisfied
    eDriftAlarm  := 3,   // 零点漂移达报警档 / Zero drift at the alarm level
    ePhaseBad    := 4    // 非法相位兜底 / Illegal phase fallback
);
END_TYPE

FUNCTION_BLOCK FB_DL_LoadCellTareDrift
VAR_INPUT
    fWeight        : REAL := 0.0;      // 当前重量读数 [kg] / Current weight reading [kg]
    bNoLoad        : BOOL := FALSE;    // 空载判定（外部给出，本件不判载荷） [-] / No-load decision, supplied externally
    fDriftWarnRate : REAL := 0.02;     // 漂移速率预警档，域 > 0.0 [kg/min] / Drift warning rate, > 0.0 [kg/min]
    fDriftAlarmRate: REAL := 0.10;     // 漂移速率报警档，域 > fDriftWarnRate [kg/min] / Drift alarm rate, > warning [kg/min]
    tObserveWin    : TIME := T#60S;    // 观测窗时长（TIME 侧），域 > T#0S [ms] / Observation window, TIME side, > 0
    fObserveWinMin : REAL := 1.0;      // 同一观测窗的分钟数值（REAL 侧），域 > eps [min] / Same window in minutes, REAL side
    fTareStableBand: REAL := 0.05;     // 去皮稳定带（|重量| 上限），域 > 0.0 [kg] / Tare stability band, > 0.0 [kg]
    tTareStable    : TIME := T#500MS;  // 去皮稳定时间，域 >= T#0S [ms] / Tare stability time, >= 0
    bTareCmd       : BOOL := FALSE;    // 去皮命令，上升沿生效 [-] / Tare command, acts on rising edge
    bReset         : BOOL := FALSE;    // 复位，上升沿清报警锁存 [-] / Reset, rising edge clears the alarm latch
END_VAR
VAR_OUTPUT
    fTareRef    : REAL;             // 当前去皮基准（零点） [kg] / Current tare reference [kg]
    fBaseline   : REAL;             // 空载基线（空载时跟随当前读数） [kg] / No-load baseline, follows the reading when empty
    fDriftRate  : REAL;             // 漂移速率（每窗末刷新，空载失效时保持） [kg/min] / Drift rate, refreshed per window
    eGrade      : E_DL_LctGrade;    // 漂移判级 [-] / Drift grade
    bTareAllowed: BOOL;             // 去皮闸放行（当拍量） [-] / Tare gate open, per scan
    bTareDone   : BOOL;             // 去皮完成，单拍脉冲 [-] / Tare done, single-scan pulse
    bTareRejected: BOOL;            // 去皮被拒（当拍量） [-] / Tare rejected
    bAlarm      : BOOL;             // 漂移报警锁存 [-] / Latched drift alarm
    eState      : E_DL_LctState;    // 状态出口 [-] / State outlet
    eCause      : E_DL_LctCause;    // 成因出口（R190 归因唯一） [-] / Cause outlet
    bError      : BOOL;             // 故障标志（组态故障或漂移报警） [-] / Error flag
END_VAR
VAR
    _eState   : E_DL_LctState := E_DL_LctState.eIdle;    // 内部相位（CASE 唯一写入目标） / Internal phase
    _eCause   : E_DL_LctCause := E_DL_LctCause.eNone;    // 成因锁存量 / Latched cause
    tonObserve: TON;            // 观测周期窗（自复位），段 0 无条件调用 / Periodic observation window, self-resetting
    tonStable : TON;            // 去皮稳定计时，段 0 无条件调用 / Tare stability timer
    rtTare    : R_TRIG;         // 去皮命令沿实例，段 0 无条件调用 / Tare command edge instance
    rtReset   : R_TRIG;         // 复位沿实例，段 0 无条件调用 / Reset edge instance
    _bFault   : BOOL;           // 报警锁存位（锁存量） / Latched alarm bit
    _bCfgBad  : BOOL;           // 组态非法当拍量 [-] / Illegal configuration this scan
    _bNonFin  : BOOL;           // 输入非有限当拍量 [-] / Non-finite input this scan
    _bStable  : BOOL;           // 空载且在稳定带内当拍量（喂稳定计时） [-] / Empty and inside the band, feeds the stability timer
    _bGate    : BOOL;           // 去皮闸当拍量 [-] / Tare gate this scan
    _bTared   : BOOL;           // 已完成过首次去皮（锁存量） / First tare done, latched
    _fRate    : REAL;           // 漂移速率锁存值（空载失效时保持） [kg/min] / Held drift rate
    _eGrade   : E_DL_LctGrade := E_DL_LctGrade.eUnknown;   // 判级锁存值（未测得时保持） / Held grade
    _fDrift   : REAL;           // 窗末漂移量中间值 [kg] / Drift at window end [kg]
END_VAR
VAR CONSTANT
    DL_LCT_EPS : REAL := 1.0E-6;    // 浮点判零容差（窗长分钟与稳定带统一口径） [无量纲] / Float epsilon
END_VAR

(* —— 段 0：当拍量派生 + 四实例无条件周期刷新 —— *)
_bNonFin := (fWeight <> fWeight) OR (fDriftWarnRate <> fDriftWarnRate)      // NaN 自反判（判等禁令唯一例外） / NaN self-reflexive tests
         OR (fDriftAlarmRate <> fDriftAlarmRate) OR (fObserveWinMin <> fObserveWinMin)
         OR (fTareStableBand <> fTareStableBand);
_bCfgBad := (tObserveWin <= T#0S) OR (fObserveWinMin <= DL_LCT_EPS)        // 窗长双口径闸（TIME 与 REAL 都要合法） / Window gates on both representations
         OR (fDriftWarnRate <= 0.0) OR (fDriftAlarmRate <= fDriftWarnRate) // 速率档几何闸 / Rate threshold geometry
         OR (fTareStableBand <= 0.0) OR (tTareStable < T#0S) OR _bNonFin;  // 稳定带与时间闸 + 非有限 / Band, time and non-finite gates
_bStable := bNoLoad AND (ABS(fWeight) <= fTareStableBand) AND (NOT _bCfgBad);   // 空载且稳定带内 / Empty and inside the stability band
_bGate   := _bStable AND tonStable.Q;                                       // 去皮闸 = 稳定且稳定时长到 / Gate = stable and duration met
rtTare(CLK := bTareCmd);                                                    // 去皮命令沿，每拍必调（R228A） / Tare edge, every scan
rtReset(CLK := bReset);                                                     // 复位沿，每拍必调 / Reset edge, every scan
tonStable(IN := _bStable, PT := tTareStable);                               // 去皮稳定计时（IN 由当拍判据派生） / Tare stability timer
tonObserve(IN := (NOT tonObserve.Q) AND bNoLoad AND (NOT _bCfgBad), PT := tObserveWin);   // 周期观测窗，自复位（R188） / Periodic window, self-resetting

(* —— 段 1：单拍量预清零（锁存量 _bFault / _fRate / _eGrade / _bTared 不入清单，R107） —— *)
bTareAllowed  := FALSE;     // 去皮闸出口每拍预清 / Gate outlet preset
bTareDone     := FALSE;     // 去皮完成每拍预清 / Tare-done pulse preset
bTareRejected := FALSE;     // 被拒标志每拍预清 / Rejected flag preset
bAlarm        := FALSE;     // 报警出口每拍预清 / Alarm outlet preset
bError        := FALSE;     // 故障标志每拍预清（R45 配对） / Error flag preset

(* —— 段 2：复位沿 + 组态闸 —— *)
IF rtReset.Q THEN
    _bFault := FALSE;                                       // 清报警锁存 / Clear alarm latch
    _eCause := E_DL_LctCause.eNone;                         // 清成因 / Clear cause
    _fRate  := 0.0;                                         // 速率锁存归零（复位即有意重开统计） / Reset the held rate deliberately
    _eGrade := E_DL_LctGrade.eUnknown;                      // 判级归未测 / Grade back to unknown
    IF _eState = E_DL_LctState.eFault THEN
        _eState := E_DL_LctState.eIdle;                     // 故障相迁出（R228B） / Leave fault phase
    END_IF
END_IF
IF _bCfgBad THEN
    _eState := E_DL_LctState.eFault;                        // 组态非法入故障相 / Enter fault phase
    _eCause := E_DL_LctCause.eCfgIllegal;                   // 归因：组态非法 / Cause: illegal configuration
END_IF

(* —— 段 3：去皮执行（命令沿 + 闸门，双条件；未放行则拒绝且不动基准） —— *)
bTareAllowed := _bGate AND (NOT _bCfgBad);                  // 闸门出口（REAL 侧与 TIME 侧均已闸） / Gate outlet
IF rtTare.Q THEN
    IF bTareAllowed THEN
        fTareRef := fWeight;                                // 取当前读数为新零点 [kg] / Present reading becomes the new zero
        fBaseline := fWeight;                               // 空载基线同步 [kg] / Baseline synchronised
        _bTared  := TRUE;                                   // 首皮完成（锁存量） / First tare done, latched
        _fRate   := 0.0;                                    // 新零点起速率重计 / Rate restarts from the new zero
        _eGrade  := E_DL_LctGrade.eOk;                      // 判级回良好 / Grade back to ok
        bTareDone := TRUE;                                  // 单拍完成脉冲 / Single-scan done pulse
    ELSE
        bTareRejected := TRUE;                              // 拒绝去皮，基准不动 / Reject, reference untouched
        _eCause := E_DL_LctCause.eTareReject;               // 归因：去皮被拒 / Cause: tare rejected
    END_IF
END_IF

(* —— 段 4：空载基线跟随（空载时基线 = 当前读数，用于 HMI 趋势） —— *)
IF bNoLoad AND (NOT _bCfgBad) THEN
    fBaseline := fWeight;                                   // 基线跟随当前读数 [kg] / Baseline follows the present reading
END_IF

(* —— 段 5：周期窗末漂移评分（单点写入 _fRate，避免同拍抹除，R187） —— *)
IF tonObserve.Q AND (NOT _bCfgBad) AND _bTared THEN
    _fDrift := fWeight - fTareRef;                          // 窗末相对去皮基准的漂移量 [kg] / Drift from the tare reference at window end
    _fRate  := _fDrift / fObserveWinMin;                    // 除以窗长分钟数得速率，分母已闸 / Rate per minute, denominator gated
    IF ABS(_fRate) >= fDriftAlarmRate THEN
        _eGrade := E_DL_LctGrade.eAlarm;                    // 报警档 / Alarm level
        _bFault := TRUE;                                    // 锁存 / Latch
        _eCause := E_DL_LctCause.eDriftAlarm;               // 归因：漂移报警 / Cause: drift alarm
    ELSIF ABS(_fRate) >= fDriftWarnRate THEN
        _eGrade := E_DL_LctGrade.eWarn;                     // 预警档（维护级，不锁存） / Warning level, maintenance only
    ELSE
        _eGrade := E_DL_LctGrade.eOk;                       // 良好档 / Ok level
    END_IF
END_IF

(* —— 段 6：锁存相位迁移闸 —— *)
IF _bFault AND (_eState <> E_DL_LctState.eFault) THEN
    _eState := E_DL_LctState.eFault;                        // 锁存即入故障相 / Latch enters fault phase
END_IF

(* —— 段 7：相位机（ENUM 全成员显式标签 + ELSE 兜底，R128） —— *)
CASE _eState OF

E_DL_LctState.eIdle:
    IF _bCfgBad THEN                                        // 出口 1：组态非法 / Illegal configuration
        _eState := E_DL_LctState.eFault;
    ELSIF _bTared THEN                                      // 出口 2：已完成去皮，进入监视 / Tare done, start monitoring
        _eState := E_DL_LctState.eRun;
    END_IF

E_DL_LctState.eRun:
    IF _bFault THEN                                         // 出口 1：漂移报警锁存 / Drift alarm latched
        _eState := E_DL_LctState.eFault;
    ELSIF (_bTared = FALSE) THEN                            // 出口 2：基准被清（复位重来） / Reference cleared, restart
        _eState := E_DL_LctState.eIdle;
    END_IF

E_DL_LctState.eFault:
    ;                                                       // 故障相：仅段 2 复位沿可迁出 / Only the reset edge leaves this phase

ELSE
    _eCause := E_DL_LctCause.ePhaseBad;                     // 归因：非法相位 / Cause: illegal phase
    _eState := E_DL_LctState.eFault;                        // 强拉故障相 / Force fault phase
    bError  := TRUE;                                        // 故障标志 / Error flag

END_CASE

(* —— 段 8：出口单点映射（名实双出口，R191） —— *)
fDriftRate := _fRate;                                       // 速率出口（空载失效时保持锁存值） / Rate outlet, held when not empty
eGrade     := _eGrade;                                      // 判级出口 / Grade outlet
bAlarm     := _bFault;                                      // 报警与锁存同源 / Alarm from latch
bError     := _bFault OR _bCfgBad;                          // 故障标志 = 锁存或组态非法 / Error = latch or illegal config
eState     := _eState;                                      // 状态出口 / State outlet
eCause     := _eCause;                                      // 成因出口 / Cause outlet

END_FUNCTION_BLOCK

(* ---- FB_DL_PdiReadScheduler.st ---- *)
(*==============================================================================
 * 组件名称 (Component)  : FB_DL_PdiReadScheduler
 * 所属子库 (Sublibrary) : DL_Device
 * 当前版本 (Version)    : 1.0.1
 * 组件分类 (Category)   : 功能块（FUNCTION_BLOCK）· 设备诊断 · 无环读取调度
 * 兼容性   (Platform)   : CODESYS 3.5 / TwinCAT 3 / 汇川 InoProShop / Schneider
 *                         Machine Expert；仅标准 TON / R_TRIG 与位运算
 * 功能描述 (Function)   : 面向参数、诊断、信息类无环读取的通用调度器。把「请求
 *                         描述域（槽、子槽、索引、子索引）加结果域（错误码、
 *                         附加信息、数据长度）」抽象成与总线无关的调度件，
 *                         硬件侧经抽象桩引脚注入就绪、完成、错误码、附加信息
 *                         与实际长度。换 RTU、换 TCP、换本地总线只换传输层，
 *                         调度层零改动。
 * 与既有件边界 (Boundary): FB_DL_ModbusPollMaster 是帧级轮询（多从站选址、
 *                         帧间静默），本件是对象字典级 PDI 调度，不触碰帧结构；
 *                         两者状态机与参数域完全不同，不得合并。
 * 工程纪律 (Discipline) : 无环通信耗时可达数十毫秒，禁止在实时任务内阻塞等待。
 *                         本块以「单拍只下发一条、忙时拒绝新启动、不排队」实现
 *                         该纪律：排队会让上层误以为指令已生效，且拖尾会累积
 *                         到下一个任务周期。
 * 设计要点 (Key notes)  : ① 请求域在启动沿一次性锁存，执行中调用方改入参不影响
 *                           在途请求；重试沿用同一锁存域，不取入参当前值；
 *                         ② 成功判据同时看错误码与数据长度：只看错误码会把
 *                           「返回长度不足」误判成功，这是无环读最常见的假成功；
 *                         ③ 失败耗尽不锁死：单次失败只记账并回待机，只有同一
 *                           请求连续三轮失败才锁故障，避免一根线缆抖动就停线；
 *                         ④ 超时用自有码（低 16 位为 5），不与总线错误码混用；
 *                         ⑤ 双层错误码打包：高 16 位附加信息、低 16 位错误码，
 *                           解包示例写在注释中，便于 HMI 直接拆。
 * 开源溯源 (Origin)     : plcnext-community。参考 PLCnext 官方公开文档所述的
 *                         无环读参数域（设备号、子设备号、对象索引、对象子索引）
 *                         与双层结果域（错误码与附加信息），以及「无环通信耗时
 *                         较长、不宜在实时任务中直接调用」的工程纪律。只借参数
 *                         域与纪律，结构体布局、状态机、码位 100% 自有
 *                         clean-room，不构成衍生作品。
 * 依赖     (Depends)    : 无 DL_ 内部依赖；仅 Standard.library 的 TON / R_TRIG
 * 故障码表 (Error codes):
 *   16#0003_013D【信息级】槽号或子槽号越界被钳位
 *   16#0003_013E【信息级】索引或子索引越界被钳位
 *   16#0003_013F【信息级】期望长度或单次超时越界被钳位
 *   16#0003_02F7【故障级】本次读取失败或超时且重试耗尽
 *   16#0003_02F8【故障级】非法状态兜底
 *   16#0003_02F9【故障级】同一请求连续三轮失败，锁定
 *   结果域自有码（写入 uErrCode 的低 16 位，不与总线码混用）：
 *   16#0000_0004 服务不可用（未使能或服务未就绪）
 *   16#0000_0005 超时
 * 验收向量 (Acceptance) :
 *   V1 成功链：服务就绪、域合法 → 启动一拍 → 请求激活 → 完成一拍且错误码 0、
 *      长度 4 → 完成脉冲单拍、成功为真、成功计数 1
 *   V2 忙时拒绝：等待期间再启动 → 拒绝计数 1、请求保持、不排队
 *   V3 重试：重试上限 1、连续两次错误码 16#0080 → 共 2 次下发后失败完成、
 *      失败计数 1、码 02F7
 *   V4 超时：不给完成信号、超时 1 秒 → 1 秒后失败完成、低 16 位为 5、
 *      请求撤回
 *   V5 打包解包：错误码 16#8011、附加信息 16#0002 → 打包值 16#0002_8011
 *   V6 长度不符：期望 8、实际 4、错误码 0 → 判失败（不得只看错误码）
 * 红线自检 (Redline)    : R1 零全局变量表与外部变量引用 ｜ R2 零物理地址直写
 *                         R3 纯 IEC 61131-3 ｜ R4 打包前显式类型转换、无浮点、
 *                         无除法 ｜ R5 全变量中英双语同行注释
 *                         R6 ENUM 加 CASE 加 ELSE 兜底 ｜ R7 TON 与两个 R_TRIG
 *                         全部在 CASE 之外无条件刷新
 * 修订历史 (Revision)   :
 *   2026-11-15  v1.0.0  首版入库（Round 10 · T1-7 PLCnext 开组）
 *   2026-11-15  v1.0.1  R10 终审修复两处：
 *                       R-FIX-1【中等】单次超时直接送进定时器 PT，未做参数域
 *                       钳位（DL_TMO_MIN / DL_TMO_MAX 两个常量声明后从未使用），
 *                       PT 填 0 会让每个等待拍立即超时形成重试风暴；补钳位并
 *                       并入 013F 参数域钳位事件（本组件码位块 013D~013F 已满，
 *                       按 R30 不得跨块取 0140，故共用 013F 并在码表说明）；
 *                       R-FIX-2【注释级】码表 013F 语义同步扩为「期望长度或
 *                       单次超时越界」。
 *============================================================================*)

(*------------------------------------------------------------------------------
 * 枚举: E_DL_PdiFsm（归属本功能块并同文件发布）
 *-----------------------------------------------------------------------------*)
TYPE E_DL_PdiFsm :
(
    eIdle  := 0,     // 待机：可受理启动沿 / Idle, accepts a start edge
    eSend  := 10,    // 下发：单拍锁存请求域并置请求激活 / Send, latches the request domain for one cycle
    eWait  := 20,    // 等待完成或超时 / Waiting for done or timeout
    eRetry := 30,    // 重试退避：单拍停留后重新下发 / Retry back-off, one cycle dwell then re-send
    eFault := 99     // 故障锁定：仅失能再使能可退 / Fault latched, only a disable-enable cycle leaves
);
END_TYPE

FUNCTION_BLOCK FB_DL_PdiReadScheduler
VAR_INPUT
    bEnable      : BOOL := TRUE;      // 使能 [-] / Enable
    bStart       : BOOL;              // 启动单次读取，上升沿；忙时忽略并计一次拒绝 [-] / Start a single read on a rising edge, ignored while busy
    uSlot        : UINT := 0;         // 设备号（槽），域 0 到 4095 [号] / Device slot number, 0 to 4095
    uSubslot     : UINT := 1;         // 子设备号（子槽），域 0 到 255 [号] / Sub-device subslot number, 0 to 255
    uIndex       : UINT := 0;         // 对象索引，域 0 到 65535 [索引] / Object index, 0 to 65535
    uSubindex    : USINT := 0;        // 对象子索引，域 0 到 255 [子索引] / Object subindex, 0 to 255
    nExpLen      : INT := 0;          // 期望数据长度，域 0 到 1024，0 表示不限 [字节] / Expected length, 0 means unrestricted
    tTimeout     : TIME := T#1S;      // 单次超时，域 100 毫秒到 10 秒 [毫秒] / Single-request timeout, 100 ms to 10 s
    nMaxRetry    : INT := 0;          // 重试次数，域 0 到 3，PDI 重试须保守 [次] / Retry count, 0 to 3, PDI retries must stay conservative
    bSrvReady    : BOOL;              // 传输层服务就绪 [-] / Transport service ready
    bSrvDone     : BOOL;              // 传输层服务完成，电平或单拍，内部取沿 [-] / Transport service done, edge detected internally
    uSrvError    : WORD;              // 服务错误码（低 16 位）[代码] / Service error code, low word of the packed result
    uSrvAddInfo  : WORD;              // 服务附加信息（高 16 位）[代码] / Service additional information, high word of the packed result
    uSrvLen      : UINT;              // 实际返回数据长度 [字节] / Actual returned data length
END_VAR
VAR_OUTPUT
    bReqActive   : BOOL;              // 请求已下发，送传输层的启动信号 [-] / Request asserted towards the transport layer
    bDone        : BOOL;              // 本次读取完成，单拍（成功或失败均置）[-] / Request finished, single-cycle pulse
    bSuccess     : BOOL;              // 本次读取成功，与完成同拍有效 [-] / TRUE when the request succeeded
    uErrCode     : UDINT;             // 双层错误码打包：高 16 位附加信息，低 16 位错误码 [代码] / Packed error code
    uActLen      : UINT;              // 实际数据长度 [字节] / Actual data length
    nRejectCnt   : UDINT;             // 忙时拒绝启动次数，跨班不清零 [次] / Busy rejection counter
    nOkCnt       : UDINT;             // 成功次数 [次] / Successful request counter
    nFailCnt     : UDINT;             // 失败次数（含重试耗尽）[次] / Failed request counter
    uErrorId     : UDINT;             // 事件码，0 = 无事件 / Event code, 0 = no event
    bError       : BOOL;              // 故障锁存，仅故障级码置位 [-] / Fault latch, set only by fault-level codes
END_VAR
VAR
    fbTrigStart  : R_TRIG;            // 启动沿检测，CASE 之外无条件刷新 [-] / Rising edge detector for the start input
    fbTrigDone   : R_TRIG;            // 完成沿检测，CASE 之外无条件刷新 [-] / Rising edge detector for the done input
    fbTmo        : TON;               // 超时计时，CASE 之外无条件刷新 [-] / Timeout timer refreshed outside the CASE
    bInit        : BOOL := FALSE;     // 首扫标志，初值 FALSE，判据 NOT bInit（R19 范式）[-] / First-scan flag
    bTmoIn       : BOOL;              // 超时定时器输入条件，先算后调以免条件调用实例 [-] / Timer input condition computed before the call
    eState       : E_DL_PdiFsm := E_DL_PdiFsm.eIdle;  // 状态机 / State machine
    nRetry       : INT;               // 本次请求已重试次数 [次] / Retries spent on the current request
    nRetryUse    : INT;               // 生效重试上限（已钳位）[次] / Effective retry limit
    nExpUse      : INT;               // 锁存的期望长度，重试沿用 [字节] / Latched expected length reused on retries
    uReqSlot     : UINT;              // 锁存的槽号 [号] / Latched slot number
    uReqSub      : UINT;              // 锁存的子槽号 [号] / Latched subslot number
    uReqIdx      : UINT;              // 锁存的索引 [索引] / Latched object index
    uReqSubIdx   : USINT;             // 锁存的子索引 [子索引] / Latched object subindex
    uSlotC       : UINT;              // 钳位后的槽号 [号] / Clamped slot number
    uSubC        : UINT;              // 钳位后的子槽号 [号] / Clamped subslot number
    nExpC        : INT;               // 钳位后的期望长度 [字节] / Clamped expected length
    tTmoUse      : TIME := T#1S;      // 钳位后的单次超时，供定时器实例使用 [毫秒] / Clamped timeout fed to the timer instance
    bOk          : BOOL;              // 本次完成的成功判据 [-] / Success predicate of the finished request
    nConsecFail  : INT;               // 同一请求连续失败轮数 [轮] / Consecutive failure rounds
    bEnablePrev  : BOOL := FALSE;     // 上拍使能值，用于失能再使能沿检测 [-] / Previous enable value for the re-enable edge
    bEnableRise  : BOOL;              // 失能再使能沿 [-] / Disable-then-enable edge
END_VAR
VAR CONSTANT
    DL_SLOT_MAX    : UINT := 4095;      // 槽号上限 [号] / Slot upper bound
    DL_SUBSLOT_MAX : UINT := 255;       // 子槽上限 [号] / Subslot upper bound
    DL_DATA_MAX    : INT  := 1024;      // 单次数据长度上限 [字节] / Data length upper bound
    DL_TMO_MIN     : TIME := T#100MS;   // 超时下限 [毫秒] / Timeout lower bound
    DL_TMO_MAX     : TIME := T#10S;     // 超时上限 [毫秒] / Timeout upper bound
    DL_RETRY_MAX   : INT  := 3;         // 重试上限，PDI 重试须保守 [次] / Retry upper bound
    DL_RETRY_MIN   : INT  := 0;         // 重试下限 [次] / Retry lower bound
    DL_FAIL_ROUNDS : INT  := 3;         // 连续失败轮数达到此值即锁故障 [轮] / Consecutive failure rounds before latching a fault
    DL_CODE_UNAVAIL: UDINT := 16#0000_0004;  // 自有码：服务不可用 [代码] / Own code, service unavailable
    DL_CODE_TIMEOUT: UDINT := 16#0000_0005;  // 自有码：超时 [代码] / Own code, timeout
    DL_PACK_SHIFT  : UDINT := 16;            // 打包移位量，附加信息移到高 16 位 [位] / Pack shift for the additional information
END_VAR

(*------------------------------------------------------------------------------
 * 段 1｜单拍输出预清零（R25 律①）
 *      Single-cycle output pre-clear
 *-----------------------------------------------------------------------------*)
bDone    := FALSE;
bSuccess := FALSE;

(*------------------------------------------------------------------------------
 * 段 2｜沿检测无条件刷新（R7 红线）
 *      Edge detection refreshed unconditionally
 *-----------------------------------------------------------------------------*)
fbTrigStart(CLK := bStart);
fbTrigDone(CLK := bSrvDone);

(*------------------------------------------------------------------------------
 * 段 3｜首扫初始化（R19 唯一合法范式）
 *      First-scan initialisation with the canonical R19 pattern
 *-----------------------------------------------------------------------------*)
IF NOT bInit THEN
    eState      := E_DL_PdiFsm.eIdle;
    nRetry      := 0;
    nConsecFail := 0;
    nOkCnt      := 0;
    nFailCnt    := 0;
    nRejectCnt  := 0;
    uErrCode    := 16#0000_0000;
    uActLen     := 0;
    bReqActive  := FALSE;
    bError      := FALSE;
    uErrorId    := 16#0000_0000;
    bInit       := TRUE;                 // 首扫只做一次
END_IF

(*------------------------------------------------------------------------------
 * 段 4｜参数域钳位（每拍，信息级）：钳位结果供启动沿锁存
 *      Parameter clamping every cycle; the start edge latches the clamped values
 *      说明：索引与子索引的取值范围由 UINT 与 USINT 类型本身饱和，越界在类型
 *      层面不可达，故 013E 分支当前为防御性保留（位宽扩展后立即生效）
 *-----------------------------------------------------------------------------*)
uSlotC := uSlot;
IF uSlotC > DL_SLOT_MAX THEN
    uSlotC  := DL_SLOT_MAX;
    uErrorId := 16#0003_013D;
END_IF

uSubC := uSubslot;
IF uSubC > DL_SUBSLOT_MAX THEN
    uSubC   := DL_SUBSLOT_MAX;
    uErrorId := 16#0003_013D;
END_IF

IF uIndex > 16#FFFF THEN
    uErrorId := 16#0003_013E;            // 防御性保留分支
END_IF
IF uSubindex > 16#FF THEN
    uErrorId := 16#0003_013E;            // 防御性保留分支
END_IF

nExpC := nExpLen;
IF nExpC < 0 THEN
    nExpC   := 0;
    uErrorId := 16#0003_013F;
ELSIF nExpC > DL_DATA_MAX THEN
    nExpC   := DL_DATA_MAX;
    uErrorId := 16#0003_013F;
END_IF

nRetryUse := nMaxRetry;
IF nRetryUse < DL_RETRY_MIN THEN
    nRetryUse := DL_RETRY_MIN;
ELSIF nRetryUse > DL_RETRY_MAX THEN
    nRetryUse := DL_RETRY_MAX;
END_IF

(* 单次超时钳位：PT 直接决定重试节奏，零或负超时会让每个等待拍立即超时，
   形成无意义的重试风暴，必须在送进定时器之前夹到合法域（红线：无魔法数、
   参数域校验）。超时钳位与期望长度钳位同属「参数域钳位」事件，共用 013F。 *)
tTmoUse := tTimeout;
IF tTmoUse < DL_TMO_MIN THEN
    tTmoUse  := DL_TMO_MIN;
    uErrorId := 16#0003_013F;
ELSIF tTmoUse > DL_TMO_MAX THEN
    tTmoUse  := DL_TMO_MAX;
    uErrorId := 16#0003_013F;
END_IF

(*------------------------------------------------------------------------------
 * 段 5｜超时计时（红线：定时器在 CASE 之外无条件刷新）
 *      Timeout timer refreshed unconditionally outside the CASE
 *-----------------------------------------------------------------------------*)
IF eState = E_DL_PdiFsm.eWait THEN
    bTmoIn := TRUE;
ELSE
    bTmoIn := FALSE;
END_IF
fbTmo(IN := bTmoIn, PT := tTmoUse);

(*------------------------------------------------------------------------------
 * 段 6｜失能再使能沿（故障态唯一退出条件）
 *      Disable-then-enable edge, the only way out of the fault state
 *-----------------------------------------------------------------------------*)
IF bEnable AND (NOT bEnablePrev) THEN
    bEnableRise := TRUE;
ELSE
    bEnableRise := FALSE;
END_IF
bEnablePrev := bEnable;

(*------------------------------------------------------------------------------
 * 段 7｜忙时拒绝计数（不排队，单拍只下发一条）
 *      Busy rejection counter, one request per cycle, never queued
 *-----------------------------------------------------------------------------*)
IF fbTrigStart.Q AND (eState <> E_DL_PdiFsm.eIdle) THEN
    nRejectCnt := nRejectCnt + 1;
END_IF

(*------------------------------------------------------------------------------
 * 段 8｜主状态机（ENUM 加 CASE，含 ELSE 兜底）
 *      Main state machine with an ELSE fallback branch
 *-----------------------------------------------------------------------------*)
CASE eState OF
    E_DL_PdiFsm.eIdle:
        bReqActive := FALSE;
        IF fbTrigStart.Q THEN
            IF (NOT bEnable) OR (NOT bSrvReady) THEN
                (* 服务不可用：立即失败完成，失败也置完成脉冲，上层才能推进 *)
                bDone       := TRUE;
                uErrCode    := DL_CODE_UNAVAIL;
                nFailCnt    := nFailCnt + 1;
                nConsecFail := nConsecFail + 1;
            ELSE
                eState := E_DL_PdiFsm.eSend;
            END_IF
        END_IF

    E_DL_PdiFsm.eSend:
        (* 单拍下发：首次下发锁存入参，重试沿用原锁存域（不取入参当前值） *)
        IF nRetry = 0 THEN
            uReqSlot   := uSlotC;
            uReqSub    := uSubC;
            uReqIdx    := uIndex;
            uReqSubIdx := uSubindex;
            nExpUse    := nExpC;
        END_IF
        bReqActive := TRUE;
        uActLen    := 0;
        eState     := E_DL_PdiFsm.eWait;

    E_DL_PdiFsm.eWait:
        bReqActive := TRUE;
        IF fbTrigDone.Q THEN
            (* 打包双层错误码：高 16 位附加信息，低 16 位错误码 *)
            uErrCode := SHL(WORD_TO_UDINT(uSrvAddInfo), DL_PACK_SHIFT) OR WORD_TO_UDINT(uSrvError);
            uActLen  := uSrvLen;
            IF (uSrvError = 16#0000) AND ((nExpUse = 0) OR (uSrvLen >= INT_TO_UINT(nExpUse))) THEN
                bOk         := TRUE;
            ELSE
                bOk         := FALSE;
            END_IF
            IF bOk THEN
                bSuccess    := TRUE;
                bDone       := TRUE;
                nOkCnt      := nOkCnt + 1;
                nConsecFail := 0;
                bReqActive  := FALSE;
                nRetry      := 0;
                eState      := E_DL_PdiFsm.eIdle;
            ELSIF nRetry < nRetryUse THEN
                nRetry     := nRetry + 1;
                bReqActive := FALSE;
                eState     := E_DL_PdiFsm.eRetry;
            ELSE
                (* 重试耗尽：本块只记账不停摆，连续三轮失败才锁故障 *)
                bDone       := TRUE;
                bSuccess    := FALSE;
                nFailCnt    := nFailCnt + 1;
                nConsecFail := nConsecFail + 1;
                bReqActive  := FALSE;
                nRetry      := 0;
                uErrorId    := 16#0003_02F7;
                IF nConsecFail >= DL_FAIL_ROUNDS THEN
                    uErrorId := 16#0003_02F9;
                    bError   := TRUE;
                    eState   := E_DL_PdiFsm.eFault;
                ELSE
                    eState := E_DL_PdiFsm.eIdle;
                END_IF
            END_IF
        ELSIF fbTmo.Q THEN
            (* 超时：撤回请求，用自有码覆盖低 16 位，再走同一重试链 *)
            bReqActive := FALSE;
            uErrCode   := DL_CODE_TIMEOUT;
            IF nRetry < nRetryUse THEN
                nRetry := nRetry + 1;
                eState := E_DL_PdiFsm.eRetry;
            ELSE
                bDone       := TRUE;
                bSuccess    := FALSE;
                nFailCnt    := nFailCnt + 1;
                nConsecFail := nConsecFail + 1;
                nRetry      := 0;
                uErrorId    := 16#0003_02F7;
                IF nConsecFail >= DL_FAIL_ROUNDS THEN
                    uErrorId := 16#0003_02F9;
                    bError   := TRUE;
                    eState   := E_DL_PdiFsm.eFault;
                ELSE
                    eState := E_DL_PdiFsm.eIdle;
                END_IF
            END_IF
        END_IF

    E_DL_PdiFsm.eRetry:
        (* 退避单拍：请求电平拉低一拍，重新下发时自然形成新的上升沿 *)
        bReqActive := FALSE;
        eState     := E_DL_PdiFsm.eSend;

    E_DL_PdiFsm.eFault:
        (* 故障锁定：请求撤回，仅失能再使能可退 *)
        bReqActive := FALSE;
        bError     := TRUE;
        IF bEnableRise THEN
            bError      := FALSE;
            uErrorId    := 16#0000_0000;
            nConsecFail := 0;
            nRetry      := 0;
            eState      := E_DL_PdiFsm.eIdle;
        END_IF

    ELSE
        (* 非法枚举值兜底 *)
        eState     := E_DL_PdiFsm.eFault;
        uErrorId   := 16#0003_02F8;
        bError     := TRUE;
        bReqActive := FALSE;
END_CASE

(*------------------------------------------------------------------------------
 * 段 9｜派生输出与解包示例（注释即文档）
 *      Derived outputs plus a worked unpacking example in comments
 *      解包示例：打包值 16#0002_8011
 *        低 16 位 = UDINT_TO_WORD(打包值 AND 16#0000_FFFF) = 16#8011（错误码）
 *        高 16 位 = UDINT_TO_WORD(SHR(打包值, 16))         = 16#0002（附加信息）
 *      注意：SHR 的移位量必须是常量或已转换的无符号量，禁止直接给有符号值
 *-----------------------------------------------------------------------------*)
IF eState = E_DL_PdiFsm.eFault THEN
    bError := TRUE;
END_IF

(*------------------------------------------------------------------------------
 * 现场提示：
 *   1 请求域在启动沿锁存后，执行期间改入参不会影响在途请求，这是刻意的：
 *     否则重试会用新参数重发，现场表现为「参数被悄悄改掉」；
 *   2 若 bSrvReady 常为假，本块只会不停返回服务不可用而不锁故障，因为这是
 *     上层联锁问题而不是本块缺陷，HMI 应把失败计数与就绪位一起显示；
 *   3 超时值不要设得比总线周期还短，否则会把「还没回」误判成「失败」，
 *     进而引发无意义的重试风暴。
 *-----------------------------------------------------------------------------*)
END_FUNCTION_BLOCK

(* ---- FB_DL_PneuCylinderDiag.st ---- *)
// ==============================================================================
// 组件名 Component  : FB_DL_PneuCylinderDiag
// 分类   Category   : DL_Device
// 前缀   Naming     : FB_DL_ ｜ b/e/t 类型前缀制（R265）
// 版本   Version    : 1.0.0
// 复杂度 Complexity  : 中
// 功能   Purpose    : 气缸纯诊断件（不控线圈）：跟踪指令沿与到位反馈的
//                      一致性——伸出 / 缩回超时（tExtTo / tRetTo）、双传感
//                      器矛盾（bFbExt 与 bFbRet 同真，物理不可能）、中途
//                      无进展（运动相中两反馈皆无持续 tStall）三族故障
//                      锁存；bReset 上升沿解锁回 eIdle。供既有气缸控制
//                      件外挂诊断层，不替代控制件。
// 开源溯源 Origin    : 道莅原创（与 FB_DL_PneumaticCylinder 的控制 + 自检
//                      一体件分工：本件为纯诊断外挂，判据独立实现
//                      clean-room，零代码复制）
// 许可证 License    : MIT
// 参考   Reference  : IEC 61131-3:2013 §6.6 ENUM + CASE 状态机 / TON /
//                      R_TRIG 语义；气缸「指令 - 反馈」一致性监视公开
//                      工程口径（借语义，不抄文）
// 平台   Platform   : 纯 IEC 61131-3（TON / R_TRIG / ENUM+CASE），三平台通用
// 依赖   Depends    : 仅 Standard.library（TON / R_TRIG 属标准件）
// 分工声明 Split     : FB_DL_PneumaticCylinder（控制件，含线圈输出与互锁）
//                      与本件互引；本件零控制出口（不下发线圈），只做
//                      指令 - 反馈一致性诊断；控制语义归彼件（R216）。
// 归属 Ownership     : E_DL_PcdSt / E_DL_PcdErr 属主为本文件（全库唯一
//                      定义，R264）；引用件只引用不重声明。
// ------------------------------------------------------------------
// 边界 Boundary     :
//   一 TON / R_TRIG 段 0 无条件刷新（禁入分支，R7）；监视 TON 串故障锁存
//      门控（FB50-1：锁存期 IN 强制 FALSE，复位同拍不重锁）；
//   二 推进判据与超时计时不同源（R300）：推进判据 = 到位反馈电平
//      （bFbExt / bFbRet），超时计时 = 状态驻留时长（tonExtTo / tonRetTo
//      基于相而非反馈），互不共源；无进展窗 tStall 为独立第三窗
//      （判据 = 两反馈皆无），与超时窗互不共源；
//   三 同拍双窗配比约束（写死）：tStall 须 < min(tExtTo, tRetTo)——
//      双反馈皆无场景下若 tStall >= 超时窗，超时窗先到，eMidStall 永不可
//      到达（配比声明，调用方改参须维持）；反馈部分在场（如 bFbRet 恒
//      真卡滞）时无进展窗被门控让路，由超时窗接管（判据互斥分层）；
//   四 故障归因唯一（R190）：eSenConflict / eMidStall / eTimeoutExt /
//      eTimeoutRet 各有独立码位与独立触发判据，禁止共用枚举成员；
//   五 eMidStall 无独立驻留相（E_DL_PcdSt 契约定稿）：锁存后冻结当前
//      运动相驻留（bErr = TRUE + eErr = eMidStall 双通道表达），迁移被
//      锁存闸（段 6）拦截至复位沿，语义在头注与码表双声明；
//   六 失败锁存 _bFaultLatch：解除式可达自证（R152）——bReset 上升沿
//      清锁存回 eIdle（输入引脚恒可达，无「置位即永久」路径）；
//   七 失能（bEn = FALSE）语义写死（R303 离相清零）：状态回 eIdle、
//      故障锁存 / 码锁存清零、bErr / bTimeout 清零（失能不是故障）；
//   八 首拍 _bInit 全量初始化（R310）；非法枚举态兜底落 eConflict +
//      eSenConflict 合并码（R90 反证句：E_DL_PcdErr 无非法态成员，非法态
//      与传感器矛盾的出口组合同为 eConflict + bErr，现有输出不可区分，
//      故合并；数值对照码 0730 见码表）；
//   九 无浮点量、无除法；无全局、无外部变量、无物理地址。
// 错误码 Codes      :
//   16#0003_0730【故障级】非法状态拦截（ELSE 兜底，经 eSenConflict 枚举
//                通道合并表达，R90 合并反证句见边界八）
//   16#0003_0731【故障级】传感器矛盾（bFbExt 与 bFbRet 同真，物理不可能）
//                → eSenConflict，锁存至复位沿
//   16#0003_0732【故障级】伸出超时（eExtending 相驻留超 tExtTo 未到位）
//                → eTimeoutExt，锁存至复位沿
//   16#0003_0733【故障级】缩回超时（eRetracting 相驻留超 tRetTo 未到位）
//                → eTimeoutRet，锁存至复位沿
//   16#0003_0734【故障级】中途无进展（运动相两反馈皆无持续 tStall）
//                → eMidStall，锁存至复位沿（冻结当前相驻留）
//   注：eErr 为枚举出口（引脚契约按任务定稿），上述数值码位为文档级
//   对照；tExtTo / tRetTo / tStall <= 0 时对应窗禁用（诊断关闭，非故障）。
// 验收 Acceptance   :
//   算法已证（脚本）：未跑 ｜ 编译器已证（三平台）：未跑
//   V1 bCmdExt 沿 + bFbExt 3s 内到位 → eExtOk、无码
//   V2 bCmdExt 沿、bFbExt 永不到 → tExtTo 到 → eExtTo + eTimeoutExt 锁存
//   V3 运动相 bFbExt 与 bFbRet 同真 → eConflict + eSenConflict 锁存
//   V4 运动相两反馈皆无超 tStall（< 超时窗）→ eMidStall 锁存、冻结驻留
//   V5 故障态 bReset 上升沿 → 解锁回 eIdle（锁存解除可达向量）
//   V6 bEn = FALSE → eIdle + 全出口清零（R303）
//   V7 非法枚举态（强改 _eState）→ ELSE 兜底落 eConflict + 0730
//   V8 tStall = T#0S → 无进展窗禁用（仅超时窗判定）
// 修订记录 Revision  :
//   2026-11-22  v1.0.0  R65 首版（批 4 · 序号 10）
// ==============================================================================
TYPE E_DL_PcdSt :
(
    eIdle       := 0,  // 空闲：等指令 / idle, waiting for the command
    eExtending  := 10, // 伸出动作中：等伸出到位反馈 / extending, waiting for the extended feedback
    eRetracting := 20, // 缩回动作中：等缩回到位反馈 / retracting, waiting for the retracted feedback
    eExtOk      := 30, // 伸出到位确认 / the extended position confirmed
    eRetOk      := 40, // 缩回到位确认 / the retracted position confirmed
    eExtTo      := 50, // 伸出超时锁存驻留（复位沿解除）/ the extend timeout dwelling, released by the reset edge
    eRetTo      := 60, // 缩回超时锁存驻留（复位沿解除）/ the retract timeout dwelling, released by the reset edge
    eConflict   := 70  // 传感器矛盾锁存驻留（复位沿解除）/ the sensor conflict dwelling, released by the reset edge
);
END_TYPE

TYPE E_DL_PcdErr :
(
    eNone        := 0,  // 无错 / no error
    eSenConflict := 10, // 传感器矛盾（含非法态拦截合并通道，边界八）/ the sensor conflict, also the illegal state channel
    eMidStall    := 20, // 中途无进展 / the mid stroke stall
    eTimeoutExt  := 30, // 伸出超时 / the extend timeout
    eTimeoutRet  := 40  // 缩回超时 / the retract timeout
);
END_TYPE

FUNCTION_BLOCK FB_DL_PneuCylinderDiag
VAR_INPUT
    bCmdExt : BOOL := FALSE;     // 伸出指令 [-]，上升沿生效 / the extend command, rising edge effective
    bCmdRet : BOOL := FALSE;     // 缩回指令 [-]，上升沿生效 / the retract command, rising edge effective
    bFbExt  : BOOL := FALSE;     // 伸出到位反馈 [-] / the extended position feedback
    bFbRet  : BOOL := FALSE;     // 缩回到位反馈 [-] / the retracted position feedback
    bEn     : BOOL := TRUE;      // 使能 [-]，FALSE 时出口清零回 eIdle（R303）/ the enable
    tExtTo  : TIME := T#5S;      // 伸出到位超时窗 [毫秒]，T#0S = 禁用 / the extend timeout, zero disables
    tRetTo  : TIME := T#5S;      // 缩回到位超时窗 [毫秒]，T#0S = 禁用 / the retract timeout, zero disables
    tStall  : TIME := T#2S;      // 无进展窗 [毫秒]，须 < min(tExtTo, tRetTo)（边界三配比），T#0S = 禁用 / the stall window with the ratio rule
    bReset  : BOOL := FALSE;     // 故障复位电平，上升沿清锁存回 eIdle（边界六解除式）/ the fault reset level
END_VAR
VAR_OUTPUT
    eSt      : E_DL_PcdSt := E_DL_PcdSt.eIdle;  // 状态机出口 [状态] / the state outlet
    bErr     : BOOL := FALSE;    // 故障锁存中 [-]，TRUE = 需复位 / the fault latched flag
    eErr     : E_DL_PcdErr := E_DL_PcdErr.eNone; // 故障码出口 [码]（锁存回放）/ the error code outlet
    bTimeout : BOOL := FALSE;    // 超时驻留指示 [-]，eExtTo / eRetTo 相为 TRUE / the timeout dwelling indicator
END_VAR
VAR
    _bInit       : BOOL := FALSE; // 首拍初始化标志（R310）/ the first scan flag
    _eState      : E_DL_PcdSt := E_DL_PcdSt.eIdle; // 内部状态寄存器 [状态] / the internal state register
    _bFaultLatch : BOOL := FALSE; // 故障锁存副本 [-]（仅复位沿清除）/ the fault latch copy
    _eErrLatch   : E_DL_PcdErr := E_DL_PcdErr.eNone; // 故障码锁存 [码]（复位沿清除，FB33-1）/ the latched error code
    rtCmdExt     : R_TRIG;        // 伸出指令沿实例，段 0 无条件刷新（R7）/ the extend command edge refreshed unconditionally
    rtCmdRet     : R_TRIG;        // 缩回指令沿实例，段 0 无条件刷新 / the retract command edge refreshed unconditionally
    rtReset      : R_TRIG;        // 复位沿实例，段 0 无条件刷新 / the reset edge instance refreshed unconditionally
    tonExtTo     : TON;           // 伸出超时窗定时器，段 0 无条件刷新 / the extend timeout timer refreshed unconditionally
    tonRetTo     : TON;           // 缩回超时窗定时器，段 0 无条件刷新 / the retract timeout timer refreshed unconditionally
    tonStall     : TON;           // 无进展窗定时器，段 0 无条件刷新 / the stall window timer refreshed unconditionally
END_VAR
VAR CONSTANT
    DL_PCD_TIME0 : TIME := T#0S; // 时间零常量 [毫秒] / the time zero constant
END_VAR

// 段 0｜定时器与沿检测实例无条件周期刷新（禁入分支，R7；监视 TON 串锁存门控，FB50-1）/ segment 0, the unconditional refresh
rtCmdExt(CLK := bCmdExt);        // 伸出指令沿 / the extend command edge
rtCmdRet(CLK := bCmdRet);        // 缩回指令沿 / the retract command edge
rtReset(CLK := bReset);          // 复位沿 / the reset edge
tonExtTo(IN := bEn AND (_eState = E_DL_PcdSt.eExtending) AND (NOT _bFaultLatch) AND (tExtTo > DL_PCD_TIME0), PT := tExtTo); // 伸出超时计时（R300：基于相驻留，与到位反馈判据不同源；窗零禁用）/ the extend timeout, state sourced per R300
tonRetTo(IN := bEn AND (_eState = E_DL_PcdSt.eRetracting) AND (NOT _bFaultLatch) AND (tRetTo > DL_PCD_TIME0), PT := tRetTo); // 缩回超时计时（同前不同源口径）/ the retract timeout, state sourced per R300
tonStall(IN := bEn AND (NOT _bFaultLatch) AND ((_eState = E_DL_PcdSt.eExtending) OR (_eState = E_DL_PcdSt.eRetracting)) AND (NOT bFbExt) AND (NOT bFbRet) AND (tStall > DL_PCD_TIME0), PT := tStall); // 无进展计时（判据 = 两反馈皆无，R300 独立第三源；反馈部分在场让路超时窗，边界三）/ the stall window on the no feedback premise

// 段 1｜首拍初始化（R310）/ segment 1, the first scan init
IF NOT _bInit THEN               // 首拍一拍 / the first scan
    _bInit := TRUE;              // 置首拍标志 / raise the first scan flag
    _eState := E_DL_PcdSt.eIdle; // 状态显式落空闲 / place the state to idle
    _bFaultLatch := FALSE;       // 故障锁存显式清零 / clear the fault latch explicitly
    _eErrLatch := E_DL_PcdErr.eNone; // 码锁存显式清零 / clear the latched code explicitly
END_IF

// 段 2｜复位沿作用域（R311：清双锁存 + 迁空闲）/ segment 2, the reset edge scope
IF rtReset.Q THEN                // 复位沿 / the reset edge
    _bFaultLatch := FALSE;       // 清故障锁存（唯一解除路径，边界六自证可达）/ clear the fault latch
    _eErrLatch := E_DL_PcdErr.eNone; // 清码锁存 / clear the latched code
    _eState := E_DL_PcdSt.eIdle; // 迁回空闲 / back to idle
END_IF

// 段 3｜失能分支：强制 eIdle + 全出口清零，不 faults（R303 离相清零声明行）/ segment 3, the disabled branch
IF NOT bEn THEN                  // 失能 / disabled
    _eState := E_DL_PcdSt.eIdle; // 强制空闲 / force the idle
    _bFaultLatch := FALSE;       // 清故障锁存（使能断开 ≠ 气缸故障）/ clear the fault latch
    _eErrLatch := E_DL_PcdErr.eNone; // 清码锁存 / clear the latched code
    eSt := _eState;              // 状态出口 / the state outlet
    bErr := FALSE;               // 故障位复位 / the fault bit resets
    eErr := E_DL_PcdErr.eNone;   // 码出口复位 / the code outlet resets
    bTimeout := FALSE;           // 超时指示复位 / the timeout indicator resets
    RETURN;                      // 早退 / early return
END_IF

// 段 4｜传感器矛盾全局闸（最高优先级，R190 归因唯一独立码；锁存期不重置）/ segment 4, the sensor conflict gate
IF bFbExt AND bFbRet AND (NOT _bFaultLatch) THEN // 双反馈同真（物理不可能，真实可达：接线错 / 磁开失效）/ both feedbacks true
    _bFaultLatch := TRUE;        // 锁存故障 / latch the fault
    _eErrLatch := E_DL_PcdErr.eSenConflict; // 故障级 0731：传感器矛盾 / the conflict code
    _eState := E_DL_PcdSt.eConflict; // 迁入矛盾驻留相 / enter the conflict phase
END_IF

// 段 5｜主状态机（ENUM + CASE + ELSE 兜底；锁存期冻结禁迁移；本拍合法事件优先于超时，R275）/ segment 5, the main machine frozen on the latch
IF NOT _bFaultLatch THEN         // 未锁存才推进（故障态 / 冻结相驻留，边界五）/ advance only without a latch
    CASE _eState OF
        E_DL_PcdSt.eIdle:        // 空闲相 / the idle phase
            IF rtCmdExt.Q THEN   // 事件优先：伸出指令沿（同拍双指令伸出优先，声明口径）/ the extend edge first
                _eState := E_DL_PcdSt.eExtending; // 迁入伸出相 / enter the extending phase
            ELSIF rtCmdRet.Q THEN // 缩回指令沿 / the retract edge
                _eState := E_DL_PcdSt.eRetracting; // 迁入缩回相 / enter the retracting phase
            END_IF
        E_DL_PcdSt.eExtending:   // 伸出相（本拍合法事件优先：到位先消化，再消化反向沿与超时窗，R275）/ the extending phase, the event before the timeout
            IF bFbExt THEN       // 到位反馈（推进判据，R300 反馈源）/ the extended feedback, the advance criterion
                _eState := E_DL_PcdSt.eExtOk; // 迁入伸出到位确认相 / enter the extended confirmed phase
            ELSIF rtCmdRet.Q THEN // 反向指令沿（中途反向合法）/ the reverse edge
                _eState := E_DL_PcdSt.eRetracting; // 迁入缩回相 / enter the retracting phase
            ELSIF tonExtTo.Q THEN // 伸出超窗（故障级 0732）/ the extend timeout
                _bFaultLatch := TRUE; // 锁存故障 / latch the fault
                _eErrLatch := E_DL_PcdErr.eTimeoutExt; // 故障码 / the extend timeout code
                _eState := E_DL_PcdSt.eExtTo; // 迁入超时驻留相 / enter the timeout dwelling phase
            ELSIF tonStall.Q THEN // 无进展超窗（故障级 0734；冻结当前相驻留，边界五）/ the stall, frozen dwelling
                _bFaultLatch := TRUE; // 锁存故障 / latch the fault
                _eErrLatch := E_DL_PcdErr.eMidStall; // 故障码 / the stall code
            END_IF               // 状态保持 eExtending（锁存闸冻结迁移，语义双声明）
        E_DL_PcdSt.eRetracting:  // 缩回相（同拍序与伸出相一致，R275）/ the retracting phase with the same event order
            IF bFbRet THEN       // 到位反馈（推进判据，R300 反馈源）/ the retracted feedback
                _eState := E_DL_PcdSt.eRetOk; // 迁入缩回到位确认相 / enter the retracted confirmed phase
            ELSIF rtCmdExt.Q THEN // 反向指令沿 / the reverse edge
                _eState := E_DL_PcdSt.eExtending; // 迁入伸出相 / enter the extending phase
            ELSIF tonRetTo.Q THEN // 缩回超窗（故障级 0733）/ the retract timeout
                _bFaultLatch := TRUE; // 锁存故障 / latch the fault
                _eErrLatch := E_DL_PcdErr.eTimeoutRet; // 故障码 / the retract timeout code
                _eState := E_DL_PcdSt.eRetTo; // 迁入超时驻留相 / enter the timeout dwelling phase
            ELSIF tonStall.Q THEN // 无进展超窗（故障级 0734；冻结当前相驻留，边界五）/ the stall, frozen dwelling
                _bFaultLatch := TRUE; // 锁存故障 / latch the fault
                _eErrLatch := E_DL_PcdErr.eMidStall; // 故障码 / the stall code
            END_IF               // 状态保持 eRetracting（锁存闸冻结迁移，语义双声明）
        E_DL_PcdSt.eExtOk:       // 伸出到位确认相（位置随反馈电平同步）/ the extended confirmed phase
            IF bFbRet AND (NOT bFbExt) THEN // 反馈切换到缩回侧 / the feedback moved to the retracted side
                _eState := E_DL_PcdSt.eRetOk; // 同步缩回确认 / sync to the retracted confirmed
            ELSIF (NOT bFbExt) AND (NOT bFbRet) THEN // 双反馈皆失（物理中途态）/ both feedbacks lost
                _eState := E_DL_PcdSt.eIdle; // 回空闲重新同步 / back to idle for a resync
            ELSIF rtCmdRet.Q THEN // 缩回指令沿 / the retract edge
                _eState := E_DL_PcdSt.eRetracting; // 迁入缩回相 / enter the retracting phase
            END_IF
        E_DL_PcdSt.eRetOk:       // 缩回到位确认相（位置随反馈电平同步）/ the retracted confirmed phase
            IF bFbExt AND (NOT bFbRet) THEN // 反馈切换到伸出侧 / the feedback moved to the extended side
                _eState := E_DL_PcdSt.eExtOk; // 同步伸出确认 / sync to the extended confirmed
            ELSIF (NOT bFbExt) AND (NOT bFbRet) THEN // 双反馈皆失 / both feedbacks lost
                _eState := E_DL_PcdSt.eIdle; // 回空闲重新同步 / back to idle for a resync
            ELSIF rtCmdExt.Q THEN // 伸出指令沿 / the extend edge
                _eState := E_DL_PcdSt.eExtending; // 迁入伸出相 / enter the extending phase
            END_IF
        E_DL_PcdSt.eExtTo:       // 伸出超时驻留相（解除由段 2 复位沿承担）/ the extend timeout dwelling, released by the reset edge
            ;                    // 驻留语义由注释表达（禁自赋值死语句，R261）/ the dwell is expressed by this comment
        E_DL_PcdSt.eRetTo:       // 缩回超时驻留相（同前驻留口径）/ the retract timeout dwelling
            ;                    // 驻留语义由注释表达 / the dwell is expressed by this comment
        E_DL_PcdSt.eConflict:    // 传感器矛盾驻留相（同前驻留口径）/ the conflict dwelling
            ;                    // 驻留语义由注释表达 / the dwell is expressed by this comment
        ELSE                     // 非法枚举值拦截（边界八：合并 eSenConflict 通道，R90 反证句见码表）/ the illegal enumeration guard
            _bFaultLatch := TRUE; // 锁存故障 / latch the fault
            _eErrLatch := E_DL_PcdErr.eSenConflict; // 故障级 0730（合并通道，R90）/ the merged conflict channel
            _eState := E_DL_PcdSt.eConflict; // 落矛盾驻留相 / force the conflict phase
    END_CASE
END_IF

// 段 6｜统一出口（名实双出口同源，R191）/ segment 6, the unified outlet
eSt := _eState;                  // 状态出口 / the state outlet
bErr := _bFaultLatch;            // 故障位与锁存同源 / the fault bit from the latch
eErr := _eErrLatch;              // 码出口与锁存同源（锁存回放）/ the code outlet from the latch
bTimeout := (_eState = E_DL_PcdSt.eExtTo) OR (_eState = E_DL_PcdSt.eRetTo); // 超时驻留指示与状态同源 / the timeout indicator from the state
END_FUNCTION_BLOCK
